(* IEC 61131-3 sources: PLC-IsaVODE/PLC-IsaVODE/samples/plc-programs (part 12) *)

(* ---- 716-TIMER_2.ST ---- *)
FUNCTION UDINT_TO_TIME2:TIME

	VAR_INPUT
		IN :	UDINT;
	END_VAR

	UDINT_TO_TIME2 := DINT_TO_TIME(UDINT_TO_DINT(IN));

END_FUNCTION

FUNCTION_BLOCK T_PLC_MS_block
	VAR_OUTPUT
		T_PLC_MS :	UDINT;
	END_VAR

	VAR_EXTERNAL
		PLC_TICKS_PER_SEC :	INT;
		PLC_SYS_TICK_CNT :	DINT;
	END_VAR

	VAR
		debug :	BOOL;(*Debug-Mode ON / OFF*)
		N :	INT;(*Debug-Faktor*)
		Offset :	UDINT;(*Debug-Offset*)
		temp :	DWORD := DWORD#1;(*Debug-Offset*)
		mode :	BOOL;(*modus*)
		faktor :	UDINT;(*Systemtakt-Faktor*)
		init :	BOOL;
		v_plc_ticks_per_sec :	UDINT;
		base :	UDINT := UDINT#1000;
	END_VAR

	IF init = FALSE THEN
		v_plc_ticks_per_sec := INT_TO_UDINT(PLC_TICKS_PER_SEC);
		IF v_plc_ticks_per_sec = UDINT#1024 THEN
			faktor := UDINT#1;
			mode := FALSE;
		ELSIF v_plc_ticks_per_sec > UDINT#0 THEN
			IF v_plc_ticks_per_sec <= base THEN
				faktor := base / v_plc_ticks_per_sec;
				mode := FALSE;
			ELSE
				faktor := v_plc_ticks_per_sec / base;
				mode := TRUE;
			END_IF;
		ELSE
			faktor := UDINT#1;
		END_IF;
		init := TRUE;
	END_IF;

	IF mode THEN
		T_PLC_MS := DINT_TO_UDINT(PLC_SYS_TICK_CNT) / faktor;
	ELSE
		T_PLC_MS := DINT_TO_UDINT(PLC_SYS_TICK_CNT) * faktor;
	END_IF;

	IF debug THEN
		T_PLC_MS := (DWORD_TO_UDINT(SHL(UDINT_TO_DWORD(T_PLC_MS),N) OR SHL(temp,N)) - UDINT#1) + Offset;
	END_IF;
END_FUNCTION_BLOCK

FUNCTION DAY_OF_WEEK:INT
  VAR_INPUT
    IDATE :	UDINT;
  END_VAR

  DAY_OF_WEEK := UDINT_TO_INT((idate / UDINT#86400 + UDINT#3) MOD UDINT#7) + INT#01;
END_FUNCTION

FUNCTION _BYTE_TO_INT:INT
	VAR_INPUT
		IN :	BYTE;
	END_VAR

	_BYTE_TO_INT := USINT_TO_INT(BYTE_TO_USINT(IN));
END_FUNCTION

FUNCTION LEAP_OF_DATE:BOOL

	VAR_INPUT
		IDATE :	UDINT;
	END_VAR

	LEAP_OF_DATE := SHL(UDINT_TO_DWORD((idate + UDINT#43200) / UDINT#31557600), 30) = DWORD#16#80000000;

END_FUNCTION

FUNCTION DAY_OF_YEAR:INT
	VAR_INPUT
		IDATE :	DATE;
	END_VAR

	DAY_OF_YEAR := UDINT_TO_INT((DATE_TO_UDINT(idate) / UDINT#86400) MOD UDINT#1461);
	IF DAY_OF_YEAR > 729 THEN
		IF DAY_OF_YEAR > 1095 THEN DAY_OF_YEAR := DAY_OF_YEAR - 1095; ELSE DAY_OF_YEAR := DAY_OF_YEAR - 729; END_IF;
	ELSIF DAY_OF_YEAR > 364 THEN
		DAY_OF_YEAR := DAY_OF_YEAR - 364;
	ELSE
		DAY_OF_YEAR := DAY_OF_YEAR + 1;
	END_IF;
END_FUNCTION

FUNCTION DAY_OF_YEAR_UDINT:INT
	VAR_INPUT
		IDATE :	UDINT;
	END_VAR

	DAY_OF_YEAR_UDINT := UDINT_TO_INT((idate / UDINT#86400) MOD UDINT#1461);
	IF DAY_OF_YEAR_UDINT > 729 THEN
		IF DAY_OF_YEAR_UDINT > 1095 THEN DAY_OF_YEAR_UDINT := DAY_OF_YEAR_UDINT - 1095; ELSE DAY_OF_YEAR_UDINT := DAY_OF_YEAR_UDINT - 729; END_IF;
	ELSIF DAY_OF_YEAR_UDINT > 364 THEN
		DAY_OF_YEAR_UDINT := DAY_OF_YEAR_UDINT - 364;
	ELSE
		DAY_OF_YEAR_UDINT := DAY_OF_YEAR_UDINT + 1;
	END_IF;
END_FUNCTION

FUNCTION MONTH_OF_DATE_UDINT:INT

	VAR_INPUT
		IDATE :	UDINT;
	END_VAR

	MONTH_OF_DATE_UDINT := DAY_OF_YEAR_UDINT(idate);
	IF MONTH_OF_DATE_UDINT < 32 THEN
		MONTH_OF_DATE_UDINT := 1;
	ELSIF LEAP_OF_DATE(IDATE) THEN
		MONTH_OF_DATE_UDINT := (MONTH_OF_DATE_UDINT * 53 + 1668) / 1623;
	ELSE
		MONTH_OF_DATE_UDINT := (MONTH_OF_DATE_UDINT * 53 + 1700) / 1620;
	END_IF;

END_FUNCTION

FUNCTION DAY_OF_MONTH:INT
	VAR_INPUT
		IDATE :	UDINT;
	END_VAR

	day_of_month := day_of_year_UDINT(idate);

	IF leap_of_Date(idate) THEN
		CASE day_of_month OF
			32..60	:	day_of_month := day_of_month - 31;
			61..91	:	day_of_month := day_of_month - 60;
			92..121 :	day_of_month := day_of_month - 91;
			122..152:	day_of_month := day_of_month - 121;
			153..182:	day_of_month := day_of_month - 152;
			183..213:	day_of_month := day_of_month - 182;
			214..244:	day_of_month := day_of_month - 213;
			245..274:	day_of_month := day_of_month - 244;
			275..305:	day_of_month := day_of_month - 274;
			306..335:	day_of_month := day_of_month - 305;
			336..366:	day_of_month := day_of_month - 335;
		END_CASE;
	ELSE
		CASE day_of_month OF
			32..59	:	day_of_month := day_of_month - 31;
			60..90	:	day_of_month := day_of_month - 59;
			91..120 :	day_of_month := day_of_month - 90;
			121..151:	day_of_month := day_of_month - 120;
			152..181:	day_of_month := day_of_month - 151;
			182..212:	day_of_month := day_of_month - 181;
			213..243:	day_of_month := day_of_month - 212;
			244..273:	day_of_month := day_of_month - 243;
			274..304:	day_of_month := day_of_month - 273;
			305..334:	day_of_month := day_of_month - 304;
			335..365:	day_of_month := day_of_month - 334;
		END_CASE;
	END_IF;

END_FUNCTION

FUNCTION MONTH_OF_DATE:INT

	VAR_INPUT
		IDATE :	DATE;
	END_VAR

	MONTH_OF_DATE := DAY_OF_YEAR(idate);
	IF MONTH_OF_DATE < 32 THEN
		MONTH_OF_DATE := 1;
	ELSIF LEAP_OF_DATE(DATE_TO_UDINT(IDATE)) THEN
		MONTH_OF_DATE := (MONTH_OF_DATE * 53 + 1668) / 1623;
	ELSE
		MONTH_OF_DATE := (MONTH_OF_DATE * 53 + 1700) / 1620;
	END_IF;

END_FUNCTION

FUNCTION TIME_TO_UDINT2:UDINT
	VAR_INPUT
		X :	TIME;
	END_VAR

	TIME_TO_UDINT2 := DINT_TO_UDINT(TIME_TO_DINT(X));
END_FUNCTION

FUNCTION DT_TO_TOD2:UDINT
	VAR_INPUT
		IN :	UDINT;
	END_VAR

	DT_TO_TOD2 := (IN MOD UDINT#86400) * UDINT#1000;
END_FUNCTION

FUNCTION _DT_TO_DATE_B:UDINT

	VAR_INPUT
		_INN :	UDINT;
	END_VAR

	_DT_TO_DATE_B := (_INN / UDINT#86400) * UDINT#86400;
END_FUNCTION

FUNCTION_BLOCK TIMER_2_Block

	VAR_INPUT
		DT_IN :	UDINT;
		START :	UDINT;
		DURATION :	TIME;
		MODE :	BYTE;
		HOLIDAY :	BOOL;
	END_VAR

	VAR_OUTPUT
		Q :	BOOL;
	END_VAR

	VAR
		last_check :	TIME := T#0s;
		dat :	UDINT;
		daytime :	UDINT;
		activation :	TIME;
		tx :	TIME;
		enabled :	BOOL;
		wday :	INT;
		init :	BOOL;
	END_VAR

	VAR RETAIN
		run_date :	UDINT;
	END_VAR

	VAR
		T_PLC_MS :	T_PLC_MS_Block;
	END_VAR

	T_PLC_MS();
	tx:= UDINT_TO_TIME(T_PLC_MS.T_PLC_MS);

	IF NOT init THEN
		init := TRUE;
		last_check := tx - t#100ms;
	END_IF;

	IF tx - last_check < T#100ms THEN RETURN; END_IF;

	dat := _DT_TO_DATE_B(dt_in);
	daytime := DT_TO_TOD2(dt_in);
	wday := DAY_OF_WEEK(dat);

	CASE _BYTE_TO_INT(mode) OF
	1..7:
		enabled := wday = _BYTE_TO_INT(mode);
	11:
		enabled := TRUE;
	12..16:
		enabled := (dat / UDINT#86400) MOD (BYTE_TO_UDINT(mode) - UDINT#10) = UDINT#0;
	20:
		enabled := wday <= 5;
	21:
		enabled := wday > 5;
	22:
		enabled := wday <= 5 AND NOT holiday;
	23:
		enabled := wday > 5 OR holiday;
	24:
		enabled := holiday;
	25:
		enabled := DAY_OF_MONTH(dat) = 1;
	26:
		enabled := day_of_month(dat + TIME_TO_UDINT2(t#1d)) = 1;
	27:
		enabled := DAY_OF_MONTH(dat) = 31 AND MONTH_OF_DATE_UDINT(dat) = 12;
	28:
		enabled := DAY_OF_YEAR_UDINT(dat) = 1;
	ELSE
		enabled := FALSE;
	END_CASE;

	IF enabled AND NOT Q AND daytime >= start AND run_date <> dat THEN
		Q := TRUE;
		activation := tx;
		run_date := dat;
	ELSIF Q AND tx - activation >= duration THEN
		Q := FALSE;
	END_IF;
	last_check := Tx;

END_FUNCTION_BLOCK

PROGRAM program0
	VAR
		DT_IN :	UDINT;
		START :	UDINT;
		DURATION :	TIME;
		MODE :	BYTE;
		HOLIDAY :	BOOL;
		Q :	BOOL;

		func_block : TIMER_2_Block;
	END_VAR
	func_block.DT_IN := DT_IN;
	func_block.START := START;
	func_block.DURATION := DURATION ;
	func_block.MODE    := MODE    ;
	func_block.HOLIDAY := HOLIDAY;

	func_block();
	Q  := func_block.Q;
END_PROGRAM

CONFIGURATION Config0
	VAR_GLOBAL
		PLC_TICKS_PER_SEC :	INT;
		PLC_SYS_TICK_CNT :	DINT;
	END_VAR
  	RESOURCE Res0 ON PLC
    	TASK task0(INTERVAL := T#20ms,PRIORITY := 0);
    	PROGRAM instance0 WITH task0 : program0;
  	END_RESOURCE
END_CONFIGURATION

(* ---- 717-SEQUENCE_8.ST ---- *)
FUNCTION UDINT_TO_TIME2:TIME

	VAR_INPUT
		IN :	UDINT;
	END_VAR

	UDINT_TO_TIME2 := DINT_TO_TIME(UDINT_TO_DINT(IN));

END_FUNCTION

FUNCTION_BLOCK T_PLC_MS_block
	VAR_OUTPUT
		T_PLC_MS :	UDINT;
	END_VAR

	VAR_EXTERNAL
		PLC_TICKS_PER_SEC :	INT;
		PLC_SYS_TICK_CNT :	DINT;
	END_VAR

	VAR
		debug :	BOOL;
		N :	INT;
		Offset :	UDINT;
		temp :	DWORD := DWORD#1;
		mode :	BOOL;
		faktor :	UDINT;
		init :	BOOL;
		v_plc_ticks_per_sec :	UDINT;
		base :	UDINT := UDINT#1000;
	END_VAR

	IF init = FALSE THEN
		v_plc_ticks_per_sec := INT_TO_UDINT(PLC_TICKS_PER_SEC);
		IF v_plc_ticks_per_sec = UDINT#1024 THEN
			faktor := UDINT#1;
			mode := FALSE;
		ELSIF v_plc_ticks_per_sec > UDINT#0 THEN
			IF v_plc_ticks_per_sec <= base THEN
				faktor := base / v_plc_ticks_per_sec;
				mode := FALSE;
			ELSE
				faktor := v_plc_ticks_per_sec / base;
				mode := TRUE;
			END_IF;
		ELSE
			faktor := UDINT#1;
		END_IF;
		init := TRUE;
	END_IF;

	IF mode THEN
		T_PLC_MS := DINT_TO_UDINT(PLC_SYS_TICK_CNT) / faktor;
	ELSE
		T_PLC_MS := DINT_TO_UDINT(PLC_SYS_TICK_CNT) * faktor;
	END_IF;

	IF debug THEN
		T_PLC_MS := (DWORD_TO_UDINT(SHL(UDINT_TO_DWORD(T_PLC_MS),N) OR SHL(temp,N)) - UDINT#1) + Offset;
	END_IF;

END_FUNCTION_BLOCK

FUNCTION_BLOCK SEQUENCE_8_Block

	VAR_INPUT
		IN0 :	BOOL := TRUE;
		IN1 :	BOOL := TRUE;
		IN2 :	BOOL := TRUE;
		IN3 :	BOOL := TRUE;
		IN4 :	BOOL := TRUE;
		IN5 :	BOOL := TRUE;
		IN6 :	BOOL := TRUE;
		IN7 :	BOOL := TRUE;
		START :	BOOL;
		RST :	BOOL;
		WAIT0 :	TIME;
		DELAY0 :	TIME;
		WAIT1 :	TIME;
		DELAY1 :	TIME;
		WAIT2 :	TIME;
		DELAY2 :	TIME;
		WAIT3 :	TIME;
		DELAY3 :	TIME;
		WAIT4 :	TIME;
		DELAY4 :	TIME;
		WAIT5 :	TIME;
		DELAY5 :	TIME;
		WAIT6 :	TIME;
		DELAY6 :	TIME;
		WAIT7 :	TIME;
		DELAY7 :	TIME;
		STOP_ON_ERROR :	BOOL;
	END_VAR

	VAR_OUTPUT
		Q0 :	BOOL;
		Q1 :	BOOL;
		Q2 :	BOOL;
		Q3 :	BOOL;
		Q4 :	BOOL;
		Q5 :	BOOL;
		Q6 :	BOOL;
		Q7 :	BOOL;
		QX :	BOOL;
		RUN :	BOOL;
		_STEP :	INT := -1;
		STATUS :	BYTE;
	END_VAR

	VAR
		last :	TIME;
		edge :	BOOL;
		tx :	TIME;
		init :	BOOL;
		T_PLC_MS :	T_PLC_MS_Block;
	END_VAR

	T_PLC_MS();
	tx:= UDINT_TO_TIME(T_PLC_MS.T_PLC_MS);

	IF NOT init THEN
		last := tx;
		init := TRUE;
		status := BYTE#110;
	END_IF;

	IF rst THEN
		_step := -1;
		Q0 := FALSE;
		Q1 := FALSE;
		Q2 := FALSE;
		Q3 := FALSE;
		Q4 := FALSE;
		Q5 := FALSE;
		Q6 := FALSE;
		Q7 := FALSE;
		status := BYTE#110;
		run := FALSE;

	ELSIF start AND NOT edge THEN
		_step := 0;
		last := tx;
		status := BYTE#111;
		Q0 := FALSE;
		Q1 := FALSE;
		Q2 := FALSE;
		Q3 := FALSE;
		Q4 := FALSE;
		Q5 := FALSE;
		Q6 := FALSE;
		Q7 := FALSE;
		run := TRUE;
	END_IF;
	edge := start;

	IF status > BYTE#0 AND status < BYTE#100 AND stop_on_error THEN RETURN; END_IF;

	IF run AND _step = 0 THEN
		IF NOT q0 AND in0 AND tx - last <= wait0 THEN
			Q0 := TRUE;
			last := tx;
		ELSIF NOT q0 AND tx - last > wait0 THEN
			status := BYTE#1;
			run := FALSE;
		ELSIF q0 AND tx - last >= delay0 THEN
			_step := 1;
			last := tx;
		END_IF;
	END_IF;
	IF run AND _step = 1 THEN
		IF NOT q1 AND in1 AND tx - last <= wait1 THEN
			Q0 := FALSE;
			Q1 := TRUE;
			last := tx;
		ELSIF NOT q1 AND Tx - last > wait1 THEN
			status := BYTE#2;
			q0 := FALSE;
			run := FALSE;
		ELSIF q1 AND tx - last >= delay1 THEN
			_step := 2;
			last := tx;
		END_IF;
	END_IF;
	IF run AND _step = 2 THEN
		IF NOT q2 AND in2 AND tx - last <= wait2 THEN
			Q1 := FALSE;
			Q2 := TRUE;
			last := tx;
		ELSIF NOT q2 AND Tx - last > wait2 THEN
			status := BYTE#3;
			q1 := FALSE;
			run := FALSE;
		ELSIF q2 AND tx - last >= delay2 THEN
			_step := 3;
			last := tx;
		END_IF;
	END_IF;
	IF run AND _step = 3 THEN
		IF NOT q3 AND in3 AND tx - last <= wait3 THEN
			Q2 := FALSE;
			Q3 := TRUE;
			last := tx;
		ELSIF NOT q3 AND Tx - last > wait3 THEN
			status := BYTE#4;
			q2 := FALSE;
			run := FALSE;
		ELSIF q3 AND tx - last >= delay3 THEN
			_step := 4;
			last := tx;
		END_IF;
	END_IF;
	IF run AND _step = 4 THEN
		IF NOT q4 AND in4 AND tx - last <= wait4 THEN
			Q3 := FALSE;
			Q4 := TRUE;
			last := tx;
		ELSIF NOT q4 AND Tx - last > wait4 THEN
			status := BYTE#5;
			q3 := FALSE;
			run := FALSE;
		ELSIF q4 AND tx - last >= delay4 THEN
			_step := 5;
			last := tx;
		END_IF;
	END_IF;
	IF run AND _step = 5 THEN
		IF NOT q5 AND in5 AND tx - last <= wait5 THEN
			Q4 := FALSE;
			Q5 := TRUE;
			last := tx;
		ELSIF NOT q5 AND Tx - last > wait5 THEN
			status := BYTE#6;
			q4 := FALSE;
			run := FALSE;
		ELSIF q5 AND tx - last >= delay5 THEN
			_step := 6;
			last := tx;
		END_IF;
	END_IF;
	IF run AND _step = 6 THEN
		IF NOT q6 AND in6 AND tx - last <= wait6 THEN
			Q5 := FALSE;
			Q6 := TRUE;
			last := tx;
		ELSIF NOT q6 AND Tx - last > wait6 THEN
			status := BYTE#7;
			q5 := FALSE;
			run := FALSE;
		ELSIF q6 AND tx - last >= delay6 THEN
			_step := 7;
			last := tx;
		END_IF;
	END_IF;
	IF run AND _step = 7 THEN
		IF NOT q7 AND in7 AND tx - last <= wait7 THEN
			Q6 := FALSE;
			Q7 := TRUE;
			last := tx;
		ELSIF NOT q7 AND Tx - last > wait7 THEN
			status := BYTE#8;
			q6 := FALSE;
			run := FALSE;
		ELSIF q7 AND tx - last >= delay7 THEN
			_step := -1;
			Q7 := FALSE;
			Run := FALSE;
			status := BYTE#110;
		END_IF;
	END_IF;
	QX := q0 OR q1 OR q2 OR q3 OR q4 OR q5 OR q6 OR q7;

END_FUNCTION_BLOCK

PROGRAM program0

	VAR
		IN0 :	BOOL := TRUE;
		IN1 :	BOOL := TRUE;
		IN2 :	BOOL := TRUE;
		IN3 :	BOOL := TRUE;
		IN4 :	BOOL := TRUE;
		IN5 :	BOOL := TRUE;
		IN6 :	BOOL := TRUE;
		IN7 :	BOOL := TRUE;
		START :	BOOL;
		RST :	BOOL;
		WAIT0 :	TIME;
		DELAY0 :	TIME;
		WAIT1 :	TIME;
		DELAY1 :	TIME;
		WAIT2 :	TIME;
		DELAY2 :	TIME;
		WAIT3 :	TIME;
		DELAY3 :	TIME;
		WAIT4 :	TIME;
		DELAY4 :	TIME;
		WAIT5 :	TIME;
		DELAY5 :	TIME;
		WAIT6 :	TIME;
		DELAY6 :	TIME;
		WAIT7 :	TIME;
		DELAY7 :	TIME;
		STOP_ON_ERROR :	BOOL;
		Q0 :	BOOL;
		Q1 :	BOOL;
		Q2 :	BOOL;
		Q3 :	BOOL;
		Q4 :	BOOL;
		Q5 :	BOOL;
		Q6 :	BOOL;
		Q7 :	BOOL;
		QX :	BOOL;
		RUN :	BOOL;
		_STEP :	INT := -1;
		STATUS :	BYTE;
		func_block : SEQUENCE_8_Block;
  	END_VAR
	func_block.IN0  :=IN0;
	func_block.IN1  :=IN1;
	func_block.IN2  :=IN2;
	func_block.IN3  :=IN3;
	func_block.IN4  :=IN4;
	func_block.IN5  :=IN5;
	func_block.IN6  :=IN6;
	func_block.IN7  :=IN7;
	func_block.START  :=START;
	func_block.RST  :=RST;
	func_block.WAIT0  :=WAIT0;
	func_block.DELAY0  :=DELAY0;
	func_block.WAIT1:=WAIT1;
	func_block.DELAY1:=DELAY1;
	func_block.WAIT2  :=WAIT2;
	func_block.DELAY2  :=DELAY2;
	func_block.WAIT3  :=WAIT3;
	func_block.DELAY3  :=DELAY3;
	func_block.DELAY1:=DELAY1;
	func_block.WAIT2  :=WAIT2;
	func_block.DELAY2  :=DELAY2;
	func_block.WAIT3  :=WAIT3;
	func_block.DELAY3  :=DELAY3;
	func_block.WAIT4:=WAIT4;
	func_block.DELAY4  :=DELAY4;
	func_block.WAIT5  :=WAIT5;
	func_block.DELAY5  :=DELAY5;
	func_block.WAIT6  :=WAIT6;
	func_block.DELAY6  :=DELAY6;
	func_block.WAIT7  :=WAIT7;
	func_block.DELAY7  :=DELAY7;
	func_block.STOP_ON_ERROR  :=STOP_ON_ERROR;
	func_block();
	Q0 := func_block.Q0;
	Q1 := func_block.Q1;
	Q2 := func_block.Q2;
	Q3 := func_block.Q3;
	Q4 := func_block.Q4;
	Q5 := func_block.Q5;
	Q6 := func_block.Q6;
	Q7 := func_block.Q7;
	QX := func_block.QX;
	RUN := func_block.RUN;
	_STEP := func_block._STEP;
	STATUS := func_block.STATUS;

END_PROGRAM

CONFIGURATION Config0

	VAR_GLOBAL
		PLC_TICKS_PER_SEC :	INT;
		PLC_SYS_TICK_CNT :	DINT;
	END_VAR

	RESOURCE Res0 ON PLC
		TASK task0(INTERVAL := T#20ms,PRIORITY := 0);
		PROGRAM instance0 WITH task0 : program0;
	END_RESOURCE

END_CONFIGURATION

(* ---- 718-BLIND_INPUT.ST ---- *)
FUNCTION UDINT_TO_TIME2:TIME

	VAR_INPUT
		IN :	UDINT;
	END_VAR

	UDINT_TO_TIME2 := DINT_TO_TIME(UDINT_TO_DINT(IN));

END_FUNCTION

FUNCTION_BLOCK T_PLC_MS_block
	VAR_OUTPUT
		T_PLC_MS :	UDINT;
	END_VAR

	VAR_EXTERNAL
		PLC_TICKS_PER_SEC :	INT;
		PLC_SYS_TICK_CNT :	DINT;
	END_VAR

	VAR
		debug :	BOOL;(*Debug-Mode ON / OFF*)
		N :	INT;(*Debug-Faktor*)
		Offset :	UDINT;(*Debug-Offset*)
		temp :	DWORD := DWORD#1;(*Debug-Offset*)
		mode :	BOOL;(*modus*)
		faktor :	UDINT;(*Systemtakt-Faktor*)
		init :	BOOL;
		v_plc_ticks_per_sec :	UDINT;
		base :	UDINT := UDINT#1000;
	END_VAR

	IF init = FALSE THEN
		v_plc_ticks_per_sec := INT_TO_UDINT(PLC_TICKS_PER_SEC);
		IF v_plc_ticks_per_sec = UDINT#1024 THEN
			faktor := UDINT#1;
			mode := FALSE;
		ELSIF v_plc_ticks_per_sec > UDINT#0 THEN
			IF v_plc_ticks_per_sec <= base THEN
				faktor := base / v_plc_ticks_per_sec;
				mode := FALSE;
			ELSE
				faktor := v_plc_ticks_per_sec / base;
				mode := TRUE;
			END_IF;
		ELSE
			faktor := UDINT#1;
		END_IF;
		init := TRUE;
	END_IF;

	IF mode THEN
		T_PLC_MS := DINT_TO_UDINT(PLC_SYS_TICK_CNT) / faktor;
	ELSE
		T_PLC_MS := DINT_TO_UDINT(PLC_SYS_TICK_CNT) * faktor;
	END_IF;

	IF debug THEN
		T_PLC_MS := (DWORD_TO_UDINT(SHL(UDINT_TO_DWORD(T_PLC_MS),N) OR SHL(temp,N)) - UDINT#1) + Offset;
	END_IF;

END_FUNCTION_BLOCK

FUNCTION_BLOCK CLICK_MODE_Block

	VAR_INPUT
		IN :	BOOL;
		T_LONG :	TIME := T#500ms;
	END_VAR

	VAR_OUTPUT
		SINGLE_ :	BOOL;
		DOUBLE :	BOOL;
		LONG :	BOOL;
		TP_LONG :	BOOL;
	END_VAR

	VAR
		Timer :	TP;
		cnt :	INT;
		last :	BOOL;
	END_VAR

	timer(in := IN, PT := T_LONG);
	single := FALSE;
	double := FALSE;

	IF timer.Q THEN
		IF NOT in AND last THEN	cnt := cnt + 1; END_IF;
	ELSE
		CASE cnt OF
			1 : single := TRUE;
			2 : double := TRUE;
		END_CASE;
		cnt := 0;
	END_IF;
	last := in;
	TP_LONG := NOT timer.Q AND (NOT LONG) AND IN;
	LONG := NOT timer.Q AND in;

END_FUNCTION_BLOCK

FUNCTION _BYTE_TO_INT:INT
	VAR_INPUT
		IN :	BYTE;
	END_VAR

	_BYTE_TO_INT := USINT_TO_INT(BYTE_TO_USINT(IN));
END_FUNCTION

FUNCTION_BLOCK BLIND_INPUT_Block

	VAR_INPUT
		POS :	BYTE;
		ANG :	BYTE;
		S1 :	BOOL;
		S2 :	BOOL;
		IN :	BOOL;
		PI :	BYTE;
		AI :	BYTE;
		SINGLE_SWITCH :	BOOL;
		CLICK_EN :	BOOL := TRUE;
		CLICK_TIME :	TIME := T#500ms;
		MAX_RUNTIME :	TIME := T#60s;
		MANUAL_TIMEOUT :	TIME := T#1h;
		DEBOUNCE_TIME :	TIME := T#20ms;
		DBL_CLK1 :	BOOL := FALSE;
		DBL_POS1 :	BYTE;
		DBL_ANG1 :	BYTE;
		DBL_CLK2 :	BOOL := FALSE;
		DBL_POS2 :	BYTE := BYTE#255;
		DBL_ANG2 :	BYTE := BYTE#255;
		D1_TOGGLE :	BOOL := TRUE;
		D2_TOGGLE :	BOOL := TRUE;
		MASTER_MODE :	BOOL;
	END_VAR

	VAR_OUTPUT
		QU :	BOOL := TRUE;
		QD :	BOOL := TRUE;
		STATUS :	BYTE;
		PO :	BYTE := BYTE#255;
		AO :	BYTE := BYTE#255;
		D1 :	BOOL;
		D2 :	BOOL;
	END_VAR

	VAR
		s1e :	TOF;
		s2e :	TOF;
		s1d :	CLICK_MODE_Block;
		s2d :	CLICK_MODE_Block;
		dir :	BOOL;
		tx :	TIME;
		last :	TIME;
		T_PLC_MS :	T_PLC_MS_Block;
	END_VAR

	T_PLC_MS();
	tx:= UDINT_TO_TIME(T_PLC_MS.T_PLC_MS);

	s1e(in := S1, pt := DEBOUNCE_TIME);
	s2e(in := S2, pt := DEBOUNCE_TIME);
	s1d(in := (s1e.Q AND NOT SINGLE_SWITCH) OR (s1e.Q AND SINGLE_SWITCH AND dir), t_long := CLICK_TIME);
	s2d(in := (s2e.Q AND NOT SINGLE_SWITCH) OR (s1e.Q AND SINGLE_SWITCH AND NOT dir), t_long := CLICK_TIME);

	IF NOT d1_toggle THEN d1 := FALSE; END_IF;
	IF NOT d2_toggle THEN d2 := FALSE; END_IF;

	IF (s1d.LONG AND s2d.LONG) OR (status = BYTE#139) THEN
	status := BYTE#139;
	IF NOT (s1d.LONG OR s2d.LONG)  THEN status := BYTE#130; END_IF;
	ELSIF s1d.tp_LONG THEN
		status := BYTE#132;
	ELSIF s2d.tp_LONG THEN
		status := BYTE#133;
	ELSIF  s1d.SINGLE_ THEN
		IF click_en THEN
			IF QU XOR QD THEN
				status := BYTE#131;
			ELSE
				status := BYTE#134;
				last := tx;
				dir := NOT dir;
			END_IF;
		END_IF;
	ELSIF  s2d.SINGLE_ THEN
		IF click_en THEN
			IF QU XOR QD THEN
				status := BYTE#131;
			ELSE
				status := BYTE#135;
				last := tx;
				dir := NOT dir;
			END_IF;
		END_IF;
	ELSIF in THEN
		status := BYTE#136;
		last := tx;
	ELSIF s1d.DOUBLE THEN
		IF dbl_clk1 THEN
			status := BYTE#137;
			last := tx;
		ELSE
			D1 := NOT D1;
		END_IF;
	ELSIF s2d.DOUBLE THEN
		IF dbl_clk2 THEN
			status := BYTE#138;
			last := tx;
		ELSE
			IF single_switch THEN D1 := NOT D1; ELSE D2 := NOT D2; END_IF;
		END_IF;
	END_IF;

	CASE _BYTE_TO_INT(status) OF
		0:
				status := BYTE#130;

		130:
				IF NOT master_mode THEN
					PO := POS;
					AO := ANG;
				END_IF;
				QU := TRUE;
				QD := TRUE;

		131:
				QU := FALSE;
				QD := FALSE;
				PO := POS;
				AO := ANG;
				IF tx - last >= manual_timeout THEN
					status := BYTE#130;
				END_IF;

		132:
				QU := TRUE;
				QD := FALSE;
				PO := POS; AO := ANG;
				last := tx;
				IF NOT s1d.LONG THEN status := BYTE#131; dir := NOT dir; END_IF;

		133:
				QU := FALSE;
				QD := TRUE;
				PO := POS; AO := ANG;
				last := tx;
				IF NOT s2d.LONG THEN	status := BYTE#131; dir := NOT dir; END_IF;

		134:
				QU := TRUE;
				QD := FALSE;
				PO := POS; AO := ANG;
				IF tx - last >= max_runtime THEN status := BYTE#131; END_IF;

		135:
				QU := FALSE;
				QD := TRUE;
				PO := POS; AO := ANG;
				IF tx - last >= max_runtime THEN status := BYTE#131;	END_IF;

		136:
				QU := TRUE;
				QD := TRUE;
				PO := PI; AO := AI;
				IF tx-last >= max_runtime THEN status := BYTE#130; END_IF;

		137:
				QU := TRUE;
				QD := TRUE;
				PO := DBL_POS1;
				AO := DBL_ANG1;
				IF tx - last >= max_runtime THEN status := BYTE#131; END_IF;

		138:
				QU := TRUE;
				QD := TRUE;
				PO := DBL_POS2;
				AO := DBL_ANG2;
				IF tx - last >= max_runtime THEN status := BYTE#131; END_IF;

		139:
				QU := FALSE;
				QD := FALSE;
				PO := POS;
				AO := ANG;

	END_CASE;

END_FUNCTION_BLOCK

PROGRAM program0
	VAR
		POS :	BYTE;
		ANG :	BYTE;
		S1 :	BOOL;
		S2 :	BOOL;
		IN :	BOOL;
		PI :	BYTE;
		AI :	BYTE;
		SINGLE_SWITCH :	BOOL;
		CLICK_EN :	BOOL := TRUE;
		CLICK_TIME :	TIME := T#500ms;
		MAX_RUNTIME :	TIME := T#60s;
		MANUAL_TIMEOUT :	TIME := T#1h;
		DEBOUNCE_TIME :	TIME := T#20ms;
		DBL_CLK1 :	BOOL := FALSE;
		DBL_POS1 :	BYTE;
		DBL_ANG1 :	BYTE;
		DBL_CLK2 :	BOOL := FALSE;
		DBL_POS2 :	BYTE := BYTE#255;
		DBL_ANG2 :	BYTE := BYTE#255;
		D1_TOGGLE :	BOOL := TRUE;
		D2_TOGGLE :	BOOL := TRUE;
		MASTER_MODE :	BOOL;
		QU :	BOOL := TRUE;
		QD :	BOOL := TRUE;
		STATUS :	BYTE;
		PO :	BYTE := BYTE#255;
		AO :	BYTE := BYTE#255;
		D1 :	BOOL;
		D2 :	BOOL;
		func_block : BLIND_INPUT_Block;
	END_VAR
	func_block.POS := POS;
	func_block.ANG := ANG;
	func_block.S1 := S1 ;
	func_block.S2 := S2;
	func_block.IN := IN;
	func_block.PI := PI;
	func_block.AI := AI;
	func_block.SINGLE_SWITCH := SINGLE_SWITCH;
	func_block.CLICK_EN := CLICK_EN ;
	func_block.CLICK_TIME := CLICK_TIME;
	func_block.MAX_RUNTIME := MAX_RUNTIME;
	func_block.MANUAL_TIMEOUT := MANUAL_TIMEOUT;
	func_block.DEBOUNCE_TIME := DEBOUNCE_TIME;
	func_block.DBL_CLK1 := DBL_CLK1;
	func_block.DBL_POS1 := DBL_POS1 ;
	func_block.DBL_ANG1 := DBL_ANG1;
	func_block.DBL_CLK2 := DBL_CLK2;
	func_block.DBL_POS2 := DBL_POS2;
	func_block.DBL_ANG2 := DBL_ANG2;
	func_block.D1_TOGGLE := D1_TOGGLE ;
	func_block.D2_TOGGLE := D2_TOGGLE;
	func_block.MASTER_MODE := MASTER_MODE;
	func_block();
	QU  := func_block.QU;
	QD  := func_block.QD;
	STATUS  := func_block.STATUS;
	PO  := func_block.PO;
	AO  := func_block.AO;
	D1  := func_block.D1;
	D2  := func_block.D2;
END_PROGRAM

CONFIGURATION Config0
	VAR_GLOBAL
		PLC_TICKS_PER_SEC :	INT;
		PLC_SYS_TICK_CNT :	DINT;
	END_VAR
  	RESOURCE Res0 ON PLC
    	TASK task0(INTERVAL := T#20ms,PRIORITY := 0);
    	PROGRAM instance0 WITH task0 : program0;
  	END_RESOURCE
END_CONFIGURATION

(* ---- 719-TN_INPUT_MENU_POPUP.ST ---- *)
FUNCTION_BLOCK TN_INPUT_MENU_POPUP

  VAR
    FB_TN_SC_AREA_SAVE :	TN_SC_AREA_SAVE;
    FB_TN_SC_AREA_RESTORE :	TN_SC_AREA_RESTORE;
    FB_TN_SC_LINE :	TN_SC_LINE;
    FB_TN_SC_ADD_SHADOW :	TN_SC_ADD_SHADOW;
    FB_TN_SC_BOX :	TN_SC_BOX;
    FB_TN_SC_WRITE_C :	TN_SC_WRITE_C;
    ELEMENT_COUNT :	ELEMENT_COUNT;
    ELEMENT_GET :	ELEMENT_GET;
  END_VAR

  VAR
    in_ROW :	INT;
    in_ROWS :	INT;
    in_COL :	INT;
    in_COLS :	INT;
    in_index :	INT;
    in_Count :	INT;
    in_Scroll_Offset :	INT;
    by_ATTR :	BYTE;
  END_VAR

  VAR_IN_OUT
    Xus_TN_MENU_POPUP :	us_TN_MENU_POPUP;
    Xus_TN_SCREEN :	us_TN_SCREEN;
  END_VAR

  IF (Xus_TN_MENU_POPUP.bo_Activ = FALSE) AND (Xus_TN_MENU_POPUP.bo_Create = TRUE) THEN
    Xus_TN_MENU_POPUP.bo_Activ         := TRUE;
    Xus_TN_MENU_POPUP.bo_Create        := FALSE;
    Xus_TN_MENU_POPUP.bo_Destroy       := FALSE;
    Xus_TN_MENU_POPUP.bo_Update        := TRUE;

    ELEMENT_COUNT(ELEMENT:=Xus_TN_MENU_POPUP.st_Menu_Text,SEP:=BYTE#35);
    Xus_TN_MENU_POPUP.st_Menu_Text:=ELEMENT_COUNT.ELEMENT;
    Xus_TN_MENU_POPUP.in_Menu_E_Count:=ELEMENT_COUNT.ELEMENT_COUNT;

    Xus_TN_MENU_POPUP.in_Rows := Xus_TN_MENU_POPUP.in_Menu_E_Count;

    Xus_TN_MENU_POPUP.in_Cols := INT#00;

    FOR in_Count := INT#01 TO Xus_TN_MENU_POPUP.in_Rows DO;

      ELEMENT_GET(ELEMENT:=Xus_TN_MENU_POPUP.st_Menu_Text,SEP:=BYTE#35,POS:=in_Count-1);
      Xus_TN_MENU_POPUP.st_Menu_Text:=ELEMENT_GET.ELEMENT;
      Xus_TN_MENU_POPUP.in_Cols:=MAX_INT(LEN(ELEMENT_GET.ELEMENT_GET),Xus_TN_MENU_POPUP.in_Cols);

    END_FOR;

    IF (Xus_TN_MENU_POPUP.in_X + Xus_TN_MENU_POPUP.in_Cols) > INT#75 THEN
      Xus_TN_MENU_POPUP.in_X := INT#79 - Xus_TN_MENU_POPUP.in_Cols - INT#04;
    END_IF;

    IF (Xus_TN_MENU_POPUP.in_Y + Xus_TN_MENU_POPUP.in_ROWS) > INT#21 THEN
      Xus_TN_MENU_POPUP.in_Y := INT#23 - Xus_TN_MENU_POPUP.in_ROWS - INT#2;
    END_IF;

    Xus_TN_SCREEN.bo_Modal_Dialog := TRUE;

    FB_TN_SC_AREA_SAVE.Iin_X1        := Xus_TN_MENU_POPUP.in_X;
    FB_TN_SC_AREA_SAVE.Iin_Y1        := Xus_TN_MENU_POPUP.in_Y;
    FB_TN_SC_AREA_SAVE.Iin_X2        := Xus_TN_MENU_POPUP.in_X + Xus_TN_MENU_POPUP.in_Cols + INT#04;
    FB_TN_SC_AREA_SAVE.Iin_Y2        := Xus_TN_MENU_POPUP.in_Y + Xus_TN_MENU_POPUP.in_Rows + INT#02;
    FB_TN_SC_AREA_SAVE.Xus_TN_SCREEN := Xus_TN_SCREEN;
    FB_TN_SC_AREA_SAVE();
    Xus_TN_SCREEN := FB_TN_SC_AREA_SAVE.Xus_TN_SCREEN;

    FB_TN_SC_BOX.Iin_X1        := Xus_TN_MENU_POPUP.in_X;
    FB_TN_SC_BOX.Iin_Y1        := Xus_TN_MENU_POPUP.in_Y;
    FB_TN_SC_BOX.Iin_X2        := Xus_TN_MENU_POPUP.in_X + Xus_TN_MENU_POPUP.in_Cols + INT#03;
    FB_TN_SC_BOX.Iin_Y2        := Xus_TN_MENU_POPUP.in_Y + Xus_TN_MENU_POPUP.in_Rows + INT#01;
    FB_TN_SC_BOX.Iby_FILL      := BYTE#32;
    FB_TN_SC_BOX.Iin_BORDER    := INT#01;
    FB_TN_SC_BOX.Iby_ATTR      := Xus_TN_MENU_POPUP.by_Attr_oF;
    FB_TN_SC_BOX.Xus_TN_SCREEN := Xus_TN_SCREEN;
    FB_TN_SC_BOX();
    Xus_TN_SCREEN := FB_TN_SC_BOX.Xus_TN_SCREEN;

    FB_TN_SC_ADD_SHADOW.Iin_X1        := Xus_TN_MENU_POPUP.in_X + INT#1;
    FB_TN_SC_ADD_SHADOW.Iin_Y1        := Xus_TN_MENU_POPUP.in_Y + INT#1;
    FB_TN_SC_ADD_SHADOW.Iin_X2        := Xus_TN_MENU_POPUP.in_X + Xus_TN_MENU_POPUP.in_Cols + INT#04;
    FB_TN_SC_ADD_SHADOW.Iin_Y2        := Xus_TN_MENU_POPUP.in_Y + Xus_TN_MENU_POPUP.in_Rows + INT#02;
    FB_TN_SC_ADD_SHADOW.Iin_OPTION    := INT#00;
    FB_TN_SC_ADD_SHADOW.Xus_TN_SCREEN := Xus_TN_SCREEN;
    FB_TN_SC_ADD_SHADOW();
    Xus_TN_SCREEN := FB_TN_SC_ADD_SHADOW.Xus_TN_SCREEN;

    in_COL  := Xus_TN_MENU_POPUP.in_X;
    in_ROW  := Xus_TN_MENU_POPUP.in_Y;
    in_ROWS := Xus_TN_MENU_POPUP.in_Rows;
    in_COLS := Xus_TN_MENU_POPUP.in_Cols;

    in_COLS := in_COLS + INT#02;

    FOR in_Count := INT#01 TO Xus_TN_MENU_POPUP.in_Menu_E_Count DO;
      in_ROW := in_ROW + INT#01;

      ELEMENT_GET(ELEMENT:=Xus_TN_MENU_POPUP.st_Menu_Text,SEP:=BYTE#35,POS:=in_Count-1);
    Xus_TN_MENU_POPUP.st_Menu_Text:=ELEMENT_GET.ELEMENT;

      IF EQ_STRING(ELEMENT_GET.ELEMENT_GET,'-') THEN

        FB_TN_SC_LINE.Iin_Y1			:= in_ROW;
        FB_TN_SC_LINE.Iin_X1			:= in_COL;
        FB_TN_SC_LINE.Iin_Y2			:= in_ROW;
        FB_TN_SC_LINE.Iin_X2			:= in_COL + in_COLS + INT#01;
        FB_TN_SC_LINE.Iby_ATTR		:= Xus_TN_MENU_POPUP.by_Attr_oF;
        FB_TN_SC_LINE.Iby_BORDER		:= BYTE#01;
        FB_TN_SC_LINE.Xus_TN_SCREEN	:= Xus_TN_SCREEN;
        FB_TN_SC_LINE();
        Xus_TN_SCREEN := FB_TN_SC_LINE.Xus_TN_SCREEN;

      END_IF;
    END_FOR;
  END_IF;

  IF (Xus_TN_MENU_POPUP.bo_Activ = TRUE) THEN

    CASE _BYTE_TO_INT(Xus_TN_MENU_POPUP.by_Input_Exten_Code) OF

    65:
      in_Scroll_Offset := INT#-1;
      Xus_TN_MENU_POPUP.bo_Update := TRUE;

    66:
      in_Scroll_Offset := INT#1;
      Xus_TN_MENU_POPUP.bo_Update := TRUE;

    13:
      Xus_TN_MENU_POPUP.bo_Destroy := TRUE;

    27:
      Xus_TN_MENU_POPUP.bo_Destroy := TRUE;
      Xus_TN_MENU_POPUP.in_Cur_Item := INT#00;

    67..68:
      Xus_TN_MENU_POPUP.bo_Destroy := TRUE;
      Xus_TN_MENU_POPUP.in_Cur_Item := INT#00;

    END_CASE;

  END_IF;

  IF (Xus_TN_MENU_POPUP.bo_Activ = TRUE) AND (Xus_TN_MENU_POPUP.bo_Update = TRUE) THEN

    Xus_TN_MENU_POPUP.bo_Update := FALSE;

    in_index := Xus_TN_MENU_POPUP.in_Cur_Item;

    IF (in_index < INT#01) OR (in_index > Xus_TN_MENU_POPUP.in_Menu_E_Count) THEN
      in_Scroll_Offset := INT#01;
      in_index := Xus_TN_MENU_POPUP.in_Menu_E_Count;
    END_IF;

    ELEMENT_GET(ELEMENT:=Xus_TN_MENU_POPUP.st_Menu_Text,SEP:=BYTE#35,POS:=in_index-1);
    Xus_TN_MENU_POPUP.st_Menu_Text:=ELEMENT_GET.ELEMENT;

    IF EQ_STRING(ELEMENT_GET.ELEMENT_GET,'-') THEN
      in_Scroll_Offset := INT#01;
    END_IF;

    IF in_Scroll_Offset <> INT#00 THEN

      FOR in_Count := INT#01 TO Xus_TN_MENU_POPUP.in_Menu_E_Count DO;

        in_index:=INC2(in_index,in_Scroll_Offset,1,Xus_TN_MENU_POPUP.in_Menu_E_Count);

        ELEMENT_GET(ELEMENT:=Xus_TN_MENU_POPUP.st_Menu_Text,SEP:=BYTE#35,POS:=in_index-1);
        Xus_TN_MENU_POPUP.st_Menu_Text:=ELEMENT_GET.ELEMENT;

        IF NE_STRING(ELEMENT_GET.ELEMENT_GET,'-') THEN
          EXIT;
        END_IF;

      END_FOR;
    END_IF;

    Xus_TN_MENU_POPUP.in_Cur_Item := in_index;
    in_Scroll_Offset := INT#00;

    in_COL  := Xus_TN_MENU_POPUP.in_X;
    in_ROW  := Xus_TN_MENU_POPUP.in_Y;
    in_ROWS := Xus_TN_MENU_POPUP.in_Rows;
    in_COLS := Xus_TN_MENU_POPUP.in_Cols;

    in_COLS := in_COLS + INT#02;

    FOR in_Count := INT#01 TO Xus_TN_MENU_POPUP.in_Menu_E_Count DO;

      in_ROW := in_ROW + INT#01;

      IF in_Count = Xus_TN_MENU_POPUP.in_Cur_Item THEN
        by_ATTR := Xus_TN_MENU_POPUP.by_Attr_mF;
      ELSE
        by_ATTR := Xus_TN_MENU_POPUP.by_Attr_oF;
      END_IF;

      ELEMENT_GET(ELEMENT:=Xus_TN_MENU_POPUP.st_Menu_Text,SEP:=BYTE#35,POS:=in_Count-1);
      Xus_TN_MENU_POPUP.st_Menu_Text:=ELEMENT_GET.ELEMENT;

      IF NE_STRING(ELEMENT_GET.ELEMENT_GET,'-') THEN

        FB_TN_SC_WRITE_C.Iin_Y         := in_ROW;
        FB_TN_SC_WRITE_C.Iin_X         := in_COL + INT#01;
        FB_TN_SC_WRITE_C.Iby_ATTR      := by_ATTR;
        FB_TN_SC_WRITE_C.Iin_LENGTH    := in_COLS;
        FB_TN_SC_WRITE_C.Iin_OPTION    := INT#02;
        FB_TN_SC_WRITE_C.Ist_STRING    := ELEMENT_GET.ELEMENT_GET;
        FB_TN_SC_WRITE_C.Xus_TN_SCREEN := Xus_TN_SCREEN;
        FB_TN_SC_WRITE_C();
        Xus_TN_SCREEN := FB_TN_SC_WRITE_C.Xus_TN_SCREEN;

      END_IF;
    END_FOR;
  END_IF;

  IF (Xus_TN_MENU_POPUP.bo_Activ = TRUE) AND (Xus_TN_MENU_POPUP.bo_Destroy = TRUE) THEN

    Xus_TN_MENU_POPUP.bo_Destroy := FALSE;
    Xus_TN_MENU_POPUP.bo_Activ   := FALSE;

    FB_TN_SC_AREA_RESTORE.Xus_TN_SCREEN := Xus_TN_SCREEN;
    FB_TN_SC_AREA_RESTORE();
    Xus_TN_SCREEN := FB_TN_SC_AREA_RESTORE.Xus_TN_SCREEN;

    Xus_TN_SCREEN.bo_Modal_Dialog := FALSE;
  END_IF;

END_FUNCTION_BLOCK

(* ---- 720-HEAT_METER.ST ---- *)
FUNCTION UDINT_TO_TIME2:TIME
	VAR_INPUT
		IN :	UDINT;
	END_VAR
	UDINT_TO_TIME2 := DINT_TO_TIME(UDINT_TO_DINT(IN));
END_FUNCTION

FUNCTION_BLOCK T_PLC_MS_block
	VAR_OUTPUT
		T_PLC_MS :	UDINT;
	END_VAR

	VAR_EXTERNAL
		PLC_TICKS_PER_SEC :	INT;
		PLC_SYS_TICK_CNT :	DINT;
	END_VAR

	VAR
		debug :	BOOL;(*Debug-Mode ON / OFF*)
		N :	INT;(*Debug-Faktor*)
		Offset :	UDINT;(*Debug-Offset*)
		temp :	DWORD := DWORD#1;(*Debug-Offset*)
		mode :	BOOL;(*modus*)
		faktor :	UDINT;(*Systemtakt-Faktor*)
		init :	BOOL;
		v_plc_ticks_per_sec :	UDINT;
		base :	UDINT := UDINT#1000;
	END_VAR

	IF init = FALSE THEN
		v_plc_ticks_per_sec := INT_TO_UDINT(PLC_TICKS_PER_SEC);
		IF v_plc_ticks_per_sec = UDINT#1024 THEN
			faktor := UDINT#1;
			mode := FALSE;
		ELSIF v_plc_ticks_per_sec > UDINT#0 THEN
			IF v_plc_ticks_per_sec <= base THEN
				faktor := base / v_plc_ticks_per_sec;
				mode := FALSE;
			ELSE
				faktor := v_plc_ticks_per_sec / base;
				mode := TRUE;
			END_IF;
		ELSE
			faktor := UDINT#1;
		END_IF;
		init := TRUE;
	END_IF;

	IF mode THEN
		T_PLC_MS := DINT_TO_UDINT(PLC_SYS_TICK_CNT) / faktor;
	ELSE
		T_PLC_MS := DINT_TO_UDINT(PLC_SYS_TICK_CNT) * faktor;
	END_IF;

	IF debug THEN
		T_PLC_MS := (DWORD_TO_UDINT(SHL(UDINT_TO_DWORD(T_PLC_MS),N) OR SHL(temp,N)) - UDINT#1) + Offset;
	END_IF;

END_FUNCTION_BLOCK

TYPE
	oscat_ARRAY_X               : ARRAY [0..1]    OF REAL;
	oscat_XY                    : ARRAY [1..20]   OF oscat_ARRAY_X := [0,0,0,0,0,0,0,0,0,0,0,0,0,0,0,0,0,0,0,0];
END_TYPE

FUNCTION_BLOCK LINEAR_INT_Block

	VAR_INPUT
		X :	REAL;
		XY :	oscat_XY;
		PTS :	INT;
	END_VAR

	VAR_OUTPUT
		LINEAR_INT :	REAL;
	END_VAR

	VAR
		i :	INT;
		i2 :	INT;
	END_VAR

	pts := MIN(pts,20);

	i := 2;

	WHILE (i < pts) AND (XY[i][0] < X) DO
		i := i + 1;
	END_WHILE;

	i2 := i-1;

	LINEAR_INT := ((XY[i][1] - XY[i2][1]) * X - XY[i][1] * XY[i2][0] + XY[i2][1] * XY[i][0]) / (XY[i][0] - XY[i2][0]);

END_FUNCTION_BLOCK

FUNCTION_BLOCK WATER_ENTHALPY_Block

    VAR_INPUT
        T :	REAL;
    END_VAR

    VAR_OUTPUT
        RESULT :	REAL;
    END_VAR

    VAR
        Pts :	INT;
        data :	oscat_XY;
        FB_LINEAR_INT :	LINEAR_INT_Block;
    END_VAR

    IF Pts = 0 THEN
        Pts := 11;
        data[01][0] := REAL#0.0;
        data[01][1] := REAL#0.06;
        data[02][0] := REAL#10.0;
        data[02][1] := REAL#42.1;
        data[03][0] := REAL#20.0;
        data[03][1] := REAL#83.9;
        data[04][0] := REAL#30.0;
        data[04][1] := REAL#125.8;
        data[05][0] := REAL#40.0;
        data[05][1] := REAL#167.58;
        data[06][0] := REAL#50.0;
        data[06][1] := REAL#209.4;
        data[07][0] := REAL#60.0;
        data[07][1] := REAL#251.2;
        data[08][0] := REAL#70.0;
        data[08][1] := REAL#293.1;
        data[09][0] := REAL#80.0;
        data[09][1] := REAL#335.0;
        data[10][0] := REAL#90.0;
        data[10][1] := REAL#377.0;
        data[11][0] := REAL#100.0;
        data[11][1] := REAL#419.1;
    END_IF;

    FB_LINEAR_INT(X:=T,XY:=Data,Pts:=Pts);
    Result :=FB_LINEAR_INT.LINEAR_INT;

END_FUNCTION_BLOCK

FUNCTION_BLOCK R2_SET_Block

	VAR_INPUT
		X :	REAL;
	END_VAR

	VAR_OUTPUT
		R2_SET :	REAL2;
	END_VAR

	R2_SET.RX := X;
	R2_SET.R1 := 0.0;

END_FUNCTION_BLOCK

FUNCTION_BLOCK R2_ADD_Block

	VAR_INPUT
		X :	REAL2;
		Y :	REAL;
	END_VAR

	VAR_OUTPUT
		R2_ADD :	REAL2;
	END_VAR

	VAR
		temp :	REAL;
	END_VAR

	temp := X.RX;
	R2_ADD.RX := Y + X.R1 + X.RX;
	R2_ADD.R1 := temp - R2_ADD.RX + Y + X.R1;

END_FUNCTION_BLOCK

TYPE REAL2:

	STRUCT
		R1 : REAL;
		RX : REAL;
	END_STRUCT;

END_TYPE

FUNCTION_BLOCK INTEGRATE

	VAR_INPUT
		E :	BOOL := TRUE;
		X :	REAL;
		K :	REAL := 1.0;
	END_VAR

	VAR_IN_OUT
		Y :	REAL;
	END_VAR

	VAR
		X_last :	REAL;
		init :	BOOL;
		T_PLC_MS :	T_PLC_MS_block;
		last :	UDINT;
		tx :	UDINT;
	END_VAR

	T_PLC_MS();
	tx:= T_PLC_MS.T_PLC_MS;

	IF NOT init THEN
		init := TRUE;
		X_last := X;
	ELSIF E THEN
		Y := (X + X_LAST) * 0.5E-3 * UDINT_TO_REAL(tx-last) * K + Y;
		X_last := X;
	END_IF;
	last := tx;

END_FUNCTION_BLOCK

FUNCTION_BLOCK FT_INT2_Block

	VAR_INPUT
		IN :	REAL;
		K :	REAL := 1.0;
		RUN :	BOOL := TRUE;
		RST :	BOOL;
		OUT_MIN :	REAL := REAL#-1.0E-37;
		OUT_MAX :	REAL := REAL#1.0E37;
	END_VAR

	VAR_OUTPUT
		OUT :	REAL;
		LIM :	BOOL;
	END_VAR

	VAR
		integ :	INTEGRATE;
		ix :	REAL;
		val :	REAL2;
		R2_ADD :	R2_ADD_Block;
		R2_SET :	R2_SET_Block;
	END_VAR

	IF RST THEN
		R2_SET(X:=0.0);
		val:=R2_SET.R2_SET;
		out := 0.0;
	ELSE
		integ(X := IN, E := RUN, K := K, Y := ix);
		ix := integ.Y;
		R2_ADD(X:=val,Y:=ix);
		val:=R2_ADD.R2_ADD;
		ix := 0.0;
		OUT := val.RX;
	END_IF;

	(* check output for limits *)
	IF out > OUT_MIN AND out < OUT_MAX THEN
		LIM := FALSE;
	ELSE
		OUT := LIMIT(OUT_MIN, OUT, OUT_MAX);
		R2_SET(X:=OUT);
		val:=R2_SET.R2_SET;
		LIM := TRUE;
	END_IF;

END_FUNCTION_BLOCK

FUNCTION WATER_DENSITY:REAL

    VAR_INPUT
        T :	REAL;
        SAT :	BOOL;
    END_VAR

    VAR
        T2 :	REAL;
        T4 :	REAL;
    END_VAR

    T2 := T * T;
    T4 := T2 * T2;
    WATER_DENSITY := (999.83952 + 16.952577*T + -7.9905127E-3*T2 + -4.6241757E-5*T2*T + 1.0584601E-7*T4 + -2.8103006E-10*T4*T) / (1.0 + 0.0168872*T);
    IF sat THEN WATER_DENSITY := WATER_DENSITY - 0.004612 + 0.000106 * T; END_IF;

END_FUNCTION

FUNCTION TIME_TO_UDINT2:UDINT
	VAR_INPUT
		X :	TIME;
	END_VAR

	TIME_TO_UDINT2 := DINT_TO_UDINT(TIME_TO_DINT(X));
END_FUNCTION

FUNCTION_BLOCK HEAT_METER_Block

	VAR_INPUT
		TF :	REAL;
		TR :	REAL;
		LPH :	REAL;
		E :	BOOL;
		RST :	BOOL;
		CP :	REAL;
		DENSITY :	REAL;
		CONTENT :	REAL;
		PULSE_MODE :	BOOL;
		RETURN_METER :	BOOL;
		AVG_TIME :	TIME := T#5s;
	END_VAR

	VAR_OUTPUT
		C :	REAL;
	END_VAR

	VAR_IN_OUT
		Y :	REAL;
	END_VAR

	VAR
		tx :	UDINT;
		last :	UDINT;
		int1 :	FT_INT2_Block;
		edge :	BOOL;
		x :	REAL;
		init :	BOOL;
		Y_last :	REAL;
		T_PLC_MS :	T_PLC_MS_Block;
		WATER_ENTHALPY :	WATER_ENTHALPY_Block;
		wa_TF :	REAL;
		wa_TR :	REAL;
	END_VAR

	IF rst THEN
		int1(rst := TRUE);
		int1.rst := FALSE;
		C := 0.0;
		Y := 0.0;
	ELSIF e THEN
		water_enthalpy(T:=TF);
		wa_TF:=water_enthalpy.Result;

		water_enthalpy(T:=TR);
		wa_TR:=water_enthalpy.Result;

		X := (WATER_DENSITY(SEL(return_meter, TF, TR), FALSE) * (wa_TF - wa_TR) * (1.0 - content) + CP * Density * content * (TF-TR));
	END_IF;

	int1(run := NOT pulse_mode AND e, in := X * LPH * 2.77777777777E-4);
	IF pulse_mode THEN
		IF NOT edge AND E THEN Y := Y + X * LPH; END_IF;
	ELSE
		Y := int1.Out;
	END_IF;

	edge := e;

	T_PLC_MS();
	tx:= T_PLC_MS.T_PLC_MS;

	IF NOT init THEN
		init := TRUE;
		last := tx;
	END_IF;

	IF (tx - last >= TIME_TO_UDINT2(AVG_TIME)) AND (avg_time > T#0s) THEN
		last := tx;
		C := (Y - Y_last) * 3.6E12 / TIME_TO_REAL(AVG_TIME);
		Y_last := Y;
	END_IF;

END_FUNCTION_BLOCK

PROGRAM program0
	VAR
	    TF :	REAL;
		TR :	REAL;
		LPH :	REAL;
		E :	BOOL;
		RST :	BOOL;
		CP :	REAL;
		DENSITY :	REAL;
		CONTENT :	REAL;
		PULSE_MODE :	BOOL;
		RETURN_METER :	BOOL;
		AVG_TIME :	TIME := T#5s;
		Y :	REAL;
		C :	REAL;

		func_block : HEAT_METER_Block;
  	END_VAR
	func_block.TF := TF;
	func_block.TR := TR;
	func_block.LPH := LPH;
	func_block.E := E;
	func_block.RST := RST;
	func_block.CP := CP;
	func_block.DENSITY := DENSITY;
	func_block.CONTENT := CONTENT;
	func_block.PULSE_MODE := PULSE_MODE;
	func_block.RETURN_METER := RETURN_METER;
	func_block.AVG_TIME := AVG_TIME;
	func_block.Y := Y;

	func_block();
	Y := func_block.Y;
	C := func_block.C;
END_PROGRAM

CONFIGURATION Config0
	VAR_GLOBAL
		PLC_TICKS_PER_SEC :	INT;
		PLC_SYS_TICK_CNT :	DINT;
	END_VAR
  	RESOURCE Res0 ON PLC
    	TASK task0(INTERVAL := T#20ms,PRIORITY := 0);
    	PROGRAM instance0 WITH task0 : program0;
  	END_RESOURCE
END_CONFIGURATION

(* ---- 721-FILE_SERVER.ST ---- *)
FUNCTION_BLOCK FILE_SERVER_Block

	VAR
		buf_size :	UDINT := UDINT#4096;
		handle :	UINT;
		read_max_length :	UDINT;
		file_position :	UDINT;
		used_filename :	STRING;
		close_time :	TIME;
		length_read :	UDINT;
		write_length :	UDINT;
		length_written :	UDINT;
		open_handle :	UINT;
		seek_mode :	UINT;
		seek_position :	UDINT;
		tell_position :	UDINT;
	END_VAR

	VAR
		last_mode :	BYTE;
		command :	BYTE;
		error_code :	BYTE;
		error :	BOOL;
		file_change :	BOOL;
		step :	INT;
		t_diff :	TIME;
		tx_last :	TIME;
		tx :	TIME;
	END_VAR

	VAR_IN_OUT
		FSD :	oscat_FILE_SERVER_DATA;
		PT :	oscat_NETWORK_BUFFER;
	END_VAR

	VAR
		FILE_REMOVE :	FILE_REMOVE;
		FILE_OPEN :	FILE_OPEN;
		FILE_SEEK :	FILE_SEEK;
		FILE_TELL :	FILE_TELL;
		FILE_CLOSE :	FILE_CLOSE;
		FILE_READ :	FILE_READ;
		FILE_WRITE :	FILE_WRITE;
		T_PLC_MS :	T_PLC_MS;
	END_VAR

	T_PLC_MS();
	tx := UDINT_TO_TIME(T_PLC_MS.T_PLC_MS);
	t_diff := tx - tx_last;
	tx_last := tx;

	CASE step OF
	0:
		IF FSD.MODE = LIMIT(BYTE#1,FSD.MODE,BYTE#5) THEN
			close_time := T#1ms;
			IF handle = UINT#00 AND FSD.MODE <= BYTE#3 THEN
				step := 100;
			ELSE
				IF EQ_STRING(used_filename, FSD.FILENAME) AND FSD.MODE = last_mode THEN
					step := 200;
				ELSE
					step := 32000;
					file_change := FSD.MODE <> BYTE#5;
				END_IF;
			END_IF;
		ELSIF handle > UINT#0 THEN
			IF FSD.AUTO_CLOSE > T#0s THEN
				close_time := close_time + t_diff;
				IF close_time > FSD.AUTO_CLOSE THEN
					step := 32000;
				END_IF;
			END_IF;
		END_IF;

	100:
		IF FSD.MODE = BYTE#3 OR FSD.MODE = BYTE#4 THEN
			command := BYTE#7;
			step := 110;
		ELSE
			step := 120;
		END_IF;

	110:
		IF command = BYTE#0  THEN
			IF (FSD.MODE = BYTE#4) OR (error and error_code <> BYTE#143) THEN
				step := 30000;
			ELSE
				step := 120;
			END_IF;
		END_IF;

	120:
		command := BYTE#1;
		last_mode := FSD.MODE;
		step := 122;

	122:
		IF command = BYTE#0 THEN
			IF error THEN
				step := 30000;
			ELSE

				close_time := T#1ms;
				handle := open_handle;
				used_filename := FSD.FILENAME;
				file_position := UDINT#4294967295;
				FSD.FILE_SIZE := UDINT#0;
				step := 125;
			END_IF;
		END_IF;

	125:
		seek_mode := UINT#2;
		seek_position := UDINT#0;
		command := BYTE#5;
		step := 130;

	130:
		IF command = BYTE#0 THEN
			IF Error THEN
				step := 30000;
			ELSE
				step := 140;
			END_IF;
		END_IF;

	140:
		command := BYTE#6;
		step := 150;

	150:
		IF command = BYTE#0 THEN
			IF Error THEN
				step := 30000;
			ELSE
				FSD.FILE_SIZE := tell_position;
				file_position := tell_position;
				FSD.FILE_OPEN := TRUE;
				step := 200;
			END_IF;
		END_IF;

	200:
		IF FSD.OFFSET > FSD.FILE_SIZE THEN
			error_code := BYTE#255;
			step := 30000;
		ELSIF FSD.OFFSET <> file_position THEN
			command := BYTE#5;
			seek_mode := UINT#0;
			seek_position := FSD.OFFSET;
			step := 210;
		ELSE
			step := 300;
		END_IF;

	210:
		IF command = BYTE#0 THEN
			file_position := seek_position;
			IF Error THEN
				step := 30000;
			ELSE
				step := 300;
			END_IF;
		END_IF;

	300:
		IF FSD.MODE = BYTE#1 THEN
			step := 400;
		ELSE
			step := 500;
		END_IF;

	400:
		IF UINT_TO_UDINT(PT.SIZE) > buf_size THEN
			read_max_length := buf_size;
		ELSE
			read_max_length := UINT_TO_UDINT(PT.SIZE);
		END_IF;

		IF file_position + read_max_length > FSD.FILE_SIZE THEN
			read_max_length := FSD.FILE_SIZE - file_position;
		END_IF;

		IF read_max_length > UDINT#0 THEN
			command := BYTE#3;
			step := INT#410;
		ELSE
			PT.SIZE := UINT#0;
			step := 30000;
		END_IF;

	410:
		IF command = BYTE#0 THEN
			PT.SIZE := UDINT_TO_UINT(length_read);
			IF NOT Error THEN
				file_position := file_position + length_read;
				FSD.OFFSET := file_position;
			END_IF;
			step := 30000;
		END_IF;

	500:
		IF UINT_TO_UDINT(PT.SIZE) > buf_size THEN
			write_length := buf_size;
		ELSE
			write_length := UINT_TO_UDINT(PT.SIZE);
		END_IF;

		IF write_length > UDINT#0 THEN
			command := BYTE#4;
			step := INT#510;
		ELSE
			step := 30000;
		END_IF;

	510:
		IF command = BYTE#0 THEN
			IF NOT Error THEN
				file_position := file_position + length_written;
				FSD.OFFSET := file_position;
				IF file_position > FSD.FILE_SIZE THEN
					FSD.FILE_SIZE := file_position;
				END_IF;
			END_IF;
			step := 30000;
		END_IF;

	30000:
		FSD.MODE := BYTE#0;
		FSD.ERROR := error_code;
		step := 0;

	32000:
		close_time := T#0s;
		IF handle > UINT#0 THEN
			command := BYTE#2;
		END_IF;
		step := 32100;

	32100:
		IF command = BYTE#0 THEN
			FSD.FILE_OPEN := FALSE;
			file_position := UDINT#0;
			FSD.FILE_SIZE := UDINT#0;
			FSD.OFFSET := UDINT#0;
			used_filename := '';
			handle := UINT#00;

			IF file_change THEN
				file_change := FALSE;
				step := 100;
			ELSE
				step := 30000;
			END_IF;
		END_IF;

	END_CASE;

	FILE_OPEN.Execute := command = BYTE#1;
	FILE_OPEN.Name := FSD.FILENAME;
	FILE_OPEN();
	open_handle := FILE_OPEN.Handle;

	IF command = BYTE#1 THEN
		IF FILE_OPEN.Done THEN
			error := FILE_OPEN.Error;
			command := BYTE#0;
			error_code := SEL_BYTE(error,BYTE#00,UINT_TO_BYTE(FILE_OPEN.ErrorID));
		END_IF;
	END_IF;

	FILE_CLOSE.Execute := command = BYTE#2;
	FILE_CLOSE.Handle := Handle;
	FILE_CLOSE();

	IF command = BYTE#2 THEN
		IF FILE_CLOSE.Done THEN
			error := FILE_CLOSE.Error;
			command := BYTE#0;
			error_code := SEL_BYTE(error,BYTE#00,UINT_TO_BYTE(FILE_CLOSE.ErrorID + UINT#10));
		END_IF;
	END_IF;

	FILE_READ.Execute := command = BYTE#3;
	FILE_READ.Handle := handle;
	FILE_READ.MaxLength := read_max_length;
	FILE_READ.Buffer := PT.BUFFER;
	FILE_READ();
	PT.BUFFER := FILE_READ.Buffer;

	IF command = BYTE#3 THEN
		IF FILE_READ.Done THEN
			error := FILE_READ.Error;
			command := BYTE#0;
			length_read :=  FILE_READ.LengthRead;
			error_code := SEL_BYTE(error,BYTE#00,UINT_TO_BYTE(FILE_READ.ErrorID + UINT#40));
		END_IF;
	END_IF;

	FILE_WRITE.Execute   := command = BYTE#4;
	FILE_WRITE.Handle    := handle;
	FILE_WRITE.Length    := write_length ;
	FILE_WRITE.Buffer    := PT.BUFFER;
	FILE_WRITE();
	PT.BUFFER := FILE_WRITE.Buffer;

	IF command = BYTE#4 THEN
		IF FILE_WRITE.Done THEN
			error := FILE_WRITE.Error;
			command := BYTE#0;
			length_written := write_length;
			error_code := SEL_BYTE(error,BYTE#00,UINT_TO_BYTE(FILE_WRITE.ErrorID + UINT#70));
		END_IF;
	END_IF;

	FILE_SEEK.Execute  := command = BYTE#5;
	FILE_SEEK.Handle   := handle;
	FILE_SEEK.Mode     := seek_mode;
	FILE_SEEK.Position := UDINT_TO_DINT(seek_position);
	FILE_SEEK();

	IF command = BYTE#5 THEN
		IF FILE_SEEK.Done THEN
			error := FILE_SEEK.Error;
			command := BYTE#0;
			error_code := SEL_BYTE(error,BYTE#00,UINT_TO_BYTE(FILE_SEEK.ErrorID + UINT#100));
		END_IF;
	END_IF;

	FILE_TELL.Execute := command = BYTE#6;
	FILE_TELL.Handle := handle;
	FILE_TELL();

	IF command = BYTE#6 THEN
		IF FILE_TELL.Done THEN
			error := FILE_TELL.Error;
			command := BYTE#0;
			tell_position := DINT_TO_UDINT(FILE_TELL.Position);
			error_code := SEL_BYTE(error,BYTE#00,UINT_TO_BYTE(FILE_TELL.ErrorID + UINT#130));
		END_IF;
	END_IF;

	FILE_REMOVE.Execute := command = BYTE#7;
	FILE_REMOVE.Name := FSD.FILENAME;
	FILE_REMOVE();

	IF command = BYTE#7 THEN
		IF FILE_REMOVE.Done THEN
			error := FILE_REMOVE.Error;
			command := BYTE#0;
			error_code := SEL_BYTE(error,BYTE#00,UINT_TO_BYTE(FILE_REMOVE.ErrorID + UINT#140));
		END_IF;
	END_IF;

END_FUNCTION_BLOCK

PROGRAM program0
	VAR
		FSD :	oscat_FILE_SERVER_DATA;
		PT :	oscat_NETWORK_BUFFER;

		func_block : FILE_SERVER_Block;
	END_VAR
	func_block.FSD := FSD;
	func_block.PT := PT;

	func_block();
	FSD  := func_block.FSD;
	PT  := func_block.PT;
END_PROGRAM

CONFIGURATION Config0
	RESOURCE Res0 ON PLC
		TASK task0(INTERVAL := T#20ms,PRIORITY := 0);
		PROGRAM instance0 WITH task0 : program0;
	END_RESOURCE
END_CONFIGURATION

(* ---- 722-BLIND_CONTROL_S.ST ---- *)
FUNCTION UDINT_TO_TIME2:TIME

	VAR_INPUT
		IN :	UDINT;
	END_VAR

	UDINT_TO_TIME2 := DINT_TO_TIME(UDINT_TO_DINT(IN));

END_FUNCTION

FUNCTION_BLOCK T_PLC_MS_block
	VAR_OUTPUT
		T_PLC_MS :	UDINT;
	END_VAR

	VAR_EXTERNAL
		PLC_TICKS_PER_SEC :	INT;
		PLC_SYS_TICK_CNT :	DINT;
	END_VAR

	VAR
		debug :	BOOL;(*Debug-Mode ON / OFF*)
		N :	INT;(*Debug-Faktor*)
		Offset :	UDINT;(*Debug-Offset*)
		temp :	DWORD := DWORD#1;(*Debug-Offset*)
		mode :	BOOL;(*modus*)
		faktor :	UDINT;(*Systemtakt-Faktor*)
		init :	BOOL;
		v_plc_ticks_per_sec :	UDINT;
		base :	UDINT := UDINT#1000;
	END_VAR

	IF init = FALSE THEN
		v_plc_ticks_per_sec := INT_TO_UDINT(PLC_TICKS_PER_SEC);
		IF v_plc_ticks_per_sec = UDINT#1024 THEN
			faktor := UDINT#1;
			mode := FALSE;
		ELSIF v_plc_ticks_per_sec > UDINT#0 THEN
			IF v_plc_ticks_per_sec <= base THEN
				faktor := base / v_plc_ticks_per_sec;
				mode := FALSE;
			ELSE
				faktor := v_plc_ticks_per_sec / base;
				mode := TRUE;
			END_IF;
		ELSE
			faktor := UDINT#1;
		END_IF;
		init := TRUE;
	END_IF;

	IF mode THEN
		T_PLC_MS := DINT_TO_UDINT(PLC_SYS_TICK_CNT) / faktor;
	ELSE
		T_PLC_MS := DINT_TO_UDINT(PLC_SYS_TICK_CNT) * faktor;
	END_IF;

	IF debug THEN
		T_PLC_MS := (DWORD_TO_UDINT(SHL(UDINT_TO_DWORD(T_PLC_MS),N) OR SHL(temp,N)) - UDINT#1) + Offset;
	END_IF;
END_FUNCTION_BLOCK

FUNCTION TIME_TO_UDINT2:UDINT
	VAR_INPUT
		X :	TIME;
	END_VAR

	TIME_TO_UDINT2 := DINT_TO_UDINT(TIME_TO_DINT(X));
END_FUNCTION

FUNCTION FRMP_B:BYTE
	VAR_INPUT
		START :	BYTE;
		DIR :	BOOL;
		TD :	TIME;
		TR :	TIME;
	END_VAR

	IF TD < TR THEN
		FRMP_B := MIN(UDINT_TO_BYTE(DWORD_TO_UDINT(SHL(TIME_TO_DWORD(TD), 8)) / TIME_TO_UDINT2(TR)), SEL(DIR, START, USINT_TO_BYTE(USINT#255 - BYTE_TO_USINT(START))));
		IF DIR THEN
			FRMP_B := USINT_TO_BYTE(BYTE_TO_USINT(START) + BYTE_TO_USINT(FRMP_B));
		ELSE
			FRMP_B := USINT_TO_BYTE(BYTE_TO_USINT(START) - BYTE_TO_USINT(FRMP_B));
		END_IF;
	ELSE
		FRMP_B := SEL(DIR, BYTE#0, BYTE#255);
	END_IF;
END_FUNCTION

FUNCTION_BLOCK _RMP_B
	VAR_INPUT
		DIR :	BOOL;
		E :	BOOL := TRUE;
		TR :	TIME;
	END_VAR

	VAR_IN_OUT
		RMP :	BYTE;
	END_VAR

	VAR
		T_PLC_MS :	T_PLC_MS_block;
		tx :	TIME;
		tl :	TIME;
		tn :	TIME;
		init :	BOOL;
		last_dir :	BOOL;
		start :	BYTE;
	END_VAR

	T_PLC_MS();
	tx := UDINT_TO_TIME(T_PLC_MS.T_PLC_MS);

	IF E AND init AND (dir = last_dir) AND (RMP <> SEL(DIR, BYTE#0, BYTE#255)) AND TR = tn THEN
		RMP := FRMP_B(start, DIR, tx - tl, TR);
	ELSE
		init := TRUE;
		tl := tx;
		tn := tr;
		start := RMP;
	END_IF;
	last_dir := dir;
END_FUNCTION_BLOCK

FUNCTION_BLOCK TREND_DW
	VAR_INPUT
		X :	DWORD;
	END_VAR
	VAR_OUTPUT
		Q :	BOOL;
		TU :	BOOL;
		TD :	BOOL;
		D :	DWORD;
	END_VAR

	VAR
		LAST_X :	DWORD;
	END_VAR

	IF X > last_X THEN
		TU := TRUE;
		TD := FALSE;
		D := UDINT_TO_DWORD(DWORD_TO_UDINT(X) - DWORD_TO_UDINT(last_X));
		Q := TRUE;
	ELSIF X < last_X THEN
		TD := TRUE;
		TU := FALSE;
		D := UDINT_TO_DWORD(DWORD_TO_UDINT(last_X) - DWORD_TO_UDINT(X));
		Q := FALSE;
	ELSE
		TU := FALSE;
		TD := FALSE;
		D := DWORD#0;
	END_IF;
	last_X := X;
END_FUNCTION_BLOCK

FUNCTION_BLOCK _RMP_NEXT
	VAR_INPUT
		E :	BOOL := TRUE;
		IN :	BYTE;
		TR :	TIME;
		TF :	TIME;
		TL :	TIME;
	END_VAR

	VAR_OUTPUT
		DIR :	BOOL;
		UP :	BOOL;
		DN :	BOOL;
	END_VAR

	VAR_IN_OUT
		OUT :	BYTE;
	END_VAR
	VAR
		rmx :	_RMP_B;
		dirx :	TREND_DW;
		t_lock :	TP;
		xen :	BOOL;
		xdir :	BOOL;
	END_VAR

	dirx(X := BYTE_TO_DWORD(in));

	t_lock(in := FALSE, pt := TL);

	IF dirx.TU AND (OUT < IN) THEN
		IF NOT xdir AND xen THEN t_lock(in := TRUE); END_IF;
		xen := TRUE;
		xdir := TRUE;
	ELSIF dirx.TD AND (OUT > IN) THEN
		IF xdir AND xen THEN t_lock(in := TRUE); END_IF;
		xen := TRUE;
		xdir := FALSE;
	ELSIF xen THEN
		IF (xdir AND (out >= in)) OR (NOT xdir AND (out <= in)) THEN
			xen := FALSE;
			IF tl > t#0s THEN t_lock(IN := TRUE); END_IF;
		END_IF;
	END_IF;

	IF NOT t_lock.Q AND xen THEN
		UP := XDIR;
		DIR := XDIR;
		DN := NOT XDIR;
	ELSE
		UP := FALSE;
		DN := FALSE;
	END_IF;

	rmx(rmp := OUT, E := E AND (UP OR DN) , dir := DIR, tr := SEL(dir, TF, TR));
	OUT := rmx.RMP;
END_FUNCTION_BLOCK

FUNCTION _BYTE_TO_INT:INT
	VAR_INPUT
		IN :	BYTE;
	END_VAR

	_BYTE_TO_INT := USINT_TO_INT(BYTE_TO_USINT(IN));
END_FUNCTION

FUNCTION_BLOCK BLIND_CONTROL_S_Block

	VAR_INPUT
		UP :	BOOL;
		DN :	BOOL;
		S_IN :	BYTE := BYTE#125;
		PI :	BYTE;
		T_UP :	TIME;
		T_DN :	TIME;
		RU :	BOOL;
		RD :	BOOL;
		T_LOCKOUT :	TIME := T#100ms;
		T_EXT :	TIME;
		EXT_TRIG :	BYTE := BYTE#5;
		R_POS_TOP :	BYTE := BYTE#255;
		R_POS_BOT :	BYTE;
	END_VAR

	VAR_OUTPUT
		POS :	BYTE;
		MU :	BOOL;
		MD :	BOOL;
		STATUS :	BYTE;
	END_VAR

	VAR
		T_PLC_MS :	T_PLC_MS_Block;
		rmp :	_RMP_NEXT;
		tx :	TIME;
		last :	TIME;
		pi_last :	BYTE;
	END_VAR

	T_PLC_MS();
	tx:= UDINT_TO_TIME(T_PLC_MS.T_PLC_MS);

	IF UP  AND NOT DN THEN
		rmp.IN := BYTE#255;
		STATUS := BYTE#121;
	ELSIF DN AND NOT UP THEN
		rmp.IN := BYTE#0;
		STATUS := BYTE#122;
	ELSIF NOT (UP OR DN) THEN
		rmp.IN := PI;
		STATUS := S_IN;
	END_IF;

	rmp(E := UP OR DN, TR := T_UP, TF := T_DN, TL := T_LOCKOUT, OUT := POS);
	pos := rmp.OUT;

	CASE _BYTE_TO_INT(STATUS) OF
		0:
			last := tx;
			PI_last := PI XOR BYTE#255;
			STATUS := BYTE#128;

		121:
			MU := TRUE;
			MD := FALSE;
			IF POS >= USINT_TO_BYTE(USINT#255 - BYTE_TO_USINT(EXT_TRIG)) THEN
				POS := BYTE#255;
				last := tx;
				STATUS := BYTE#129;
			END_IF;

		122:
			MD := TRUE;
			MU := FALSE;
			IF POS <= EXT_TRIG THEN
				POS := BYTE#0;
				last := tx;
				STATUS := BYTE#129;
			END_IF;

		123:
			MD := rmp.DN;
			MU := rmp.UP;
			IF NOT (rmp.DN OR rmp.UP) THEN
				IF POS <= EXT_TRIG THEN
					MD := TRUE;
					last := tx;
					STATUS := BYTE#129;
				ELSIF POS >= USINT_TO_BYTE(USINT#255 - BYTE_TO_USINT(EXT_TRIG)) THEN
					MU := TRUE;
					last := tx;
					STATUS := BYTE#129;
				ELSE
					STATUS := S_IN;
				END_IF;
			END_IF;

		124:
			MD := rmp.DN;
			MU := rmp.UP;
			IF NOT(rmp.DN OR rmp.UP) THEN
				PI_last := PI;
				STATUS := S_IN;
			END_IF;

		127:
			IF (tx - last) >= T_LOCKOUT THEN
					STATUS := S_IN;
			END_IF;

		128:
			MU := TRUE;
			MD := FALSE;
			rmp.IN := BYTE#255;
			IF (tx - last) >= (T_UP +  T_EXT) THEN
				MU := FALSE;
				last := tx;
				STATUS := BYTE#127;
			END_IF;

		129:
			IF (tx - last) >= T_EXT THEN
				MU := FALSE;
				MD := FALSE;
				last := tx;
				STATUS := BYTE#127;
			END_IF;

	ELSE
		MU := FALSE;
		MD := FALSE;
		IF PI <> PI_last THEN
			PI_last := PI;
			rmp.IN := PI;
			STATUS := BYTE#123;
		ELSIF POS = BYTE#0 AND RU THEN
			rmp.IN := R_POS_BOT;
			STATUS := BYTE#124;
		ELSIF pos = BYTE#255 AND RD THEN
			rmp.IN := R_POS_TOP;
			STATUS := BYTE#124;
		ELSE
			STATUS := S_IN;
		END_IF;
	END_CASE;

END_FUNCTION_BLOCK

PROGRAM program0
	VAR
		UP :	BOOL;
		DN :	BOOL;
		S_IN :	BYTE := BYTE#125;
		PI :	BYTE;
		T_UP :	TIME;
		T_DN :	TIME;
		RU :	BOOL;
		RD :	BOOL;
		T_LOCKOUT :	TIME := T#100ms;
		T_EXT :	TIME;
		EXT_TRIG :	BYTE := BYTE#5;
		R_POS_TOP :	BYTE := BYTE#255;
		R_POS_BOT :	BYTE;
		POS :	BYTE;
		MU :	BOOL;
		MD :	BOOL;
		STATUS :	BYTE;
		func_block : BLIND_CONTROL_S_Block;
	END_VAR
	func_block.UP := UP;
	func_block.DN := DN;
	func_block.S_IN := S_IN ;
	func_block.PI    := PI    ;
	func_block.T_UP := T_UP;
	func_block.T_DN := T_DN ;
	func_block.RU    := RU    ;
	func_block.RD := RD;
	func_block.T_LOCKOUT := T_LOCKOUT;
	func_block.T_EXT := T_EXT ;
	func_block.EXT_TRIG    := EXT_TRIG    ;
	func_block.R_POS_TOP := R_POS_TOP;
	func_block.R_POS_BOT := R_POS_BOT ;
	func_block();
	POS  := func_block.POS;
	MU  := func_block.MU;
	MD  := func_block.MD;
	STATUS  := func_block.STATUS;
END_PROGRAM

CONFIGURATION Config0
	VAR_GLOBAL
		PLC_TICKS_PER_SEC :	INT;
		PLC_SYS_TICK_CNT :	DINT;
	END_VAR
  	RESOURCE Res0 ON PLC
    	TASK task0(INTERVAL := T#20ms,PRIORITY := 0);
    	PROGRAM instance0 WITH task0 : program0;
  	END_RESOURCE
END_CONFIGURATION

(* ---- 723-ACTUATOR_3P.ST ---- *)
FUNCTION UDINT_TO_TIME2:TIME

	VAR_INPUT
		IN :	UDINT;
	END_VAR

	UDINT_TO_TIME2 := DINT_TO_TIME(UDINT_TO_DINT(IN));

END_FUNCTION

FUNCTION_BLOCK T_PLC_MS_block
	VAR_OUTPUT
		T_PLC_MS :	UDINT;
	END_VAR

	VAR_EXTERNAL
		PLC_TICKS_PER_SEC :	INT;
		PLC_SYS_TICK_CNT :	DINT;
	END_VAR

	VAR
		debug :	BOOL;(*Debug-Mode ON / OFF*)
		N :	INT;(*Debug-Faktor*)
		Offset :	UDINT;(*Debug-Offset*)
		temp :	DWORD := DWORD#1;(*Debug-Offset*)
		mode :	BOOL;(*modus*)
		faktor :	UDINT;(*Systemtakt-Faktor*)
		init :	BOOL;
		v_plc_ticks_per_sec :	UDINT;
		base :	UDINT := UDINT#1000;
	END_VAR

	IF init = FALSE THEN
		v_plc_ticks_per_sec := INT_TO_UDINT(PLC_TICKS_PER_SEC);
		IF v_plc_ticks_per_sec = UDINT#1024 THEN
			faktor := UDINT#1;
			mode := FALSE;
		ELSIF v_plc_ticks_per_sec > UDINT#0 THEN
			IF v_plc_ticks_per_sec <= base THEN
				faktor := base / v_plc_ticks_per_sec;
				mode := FALSE;
			ELSE
				faktor := v_plc_ticks_per_sec / base;
				mode := TRUE;
			END_IF;
		ELSE
			faktor := UDINT#1;
		END_IF;
		init := TRUE;
	END_IF;

	IF mode THEN
		T_PLC_MS := DINT_TO_UDINT(PLC_SYS_TICK_CNT) / faktor;
	ELSE
		T_PLC_MS := DINT_TO_UDINT(PLC_SYS_TICK_CNT) * faktor;
	END_IF;

	IF debug THEN
		T_PLC_MS := (DWORD_TO_UDINT(SHL(UDINT_TO_DWORD(T_PLC_MS),N) OR SHL(temp,N)) - UDINT#1) + Offset;
	END_IF;
END_FUNCTION_BLOCK

FUNCTION TIME_TO_UDINT2:UDINT
	VAR_INPUT
		X :	TIME;
	END_VAR

	TIME_TO_UDINT2 := DINT_TO_UDINT(TIME_TO_DINT(X));
END_FUNCTION

FUNCTION FRMP_B:BYTE
	VAR_INPUT
		START :	BYTE;
		DIR :	BOOL;
		TD :	TIME;
		TR :	TIME;
	END_VAR

	IF TD < TR THEN
		FRMP_B := MIN(UDINT_TO_BYTE(DWORD_TO_UDINT(SHL(TIME_TO_DWORD(TD), 8)) / TIME_TO_UDINT2(TR)), SEL(DIR, START, USINT_TO_BYTE(USINT#255 - BYTE_TO_USINT(START))));
		IF DIR THEN
			FRMP_B := USINT_TO_BYTE(BYTE_TO_USINT(START) + BYTE_TO_USINT(FRMP_B));
		ELSE
			FRMP_B := USINT_TO_BYTE(BYTE_TO_USINT(START) - BYTE_TO_USINT(FRMP_B));
		END_IF;
	ELSE
		FRMP_B := SEL(DIR, BYTE#0, BYTE#255);
	END_IF;
END_FUNCTION

FUNCTION_BLOCK _RMP_B
	VAR_INPUT
		DIR :	BOOL;
		E :	BOOL := TRUE;
		TR :	TIME;
	END_VAR

	VAR_IN_OUT
		RMP :	BYTE;
	END_VAR

	VAR
		T_PLC_MS :	T_PLC_MS_block;
		tx :	TIME;
		tl :	TIME;
		tn :	TIME;
		init :	BOOL;
		last_dir :	BOOL;
		start :	BYTE;
	END_VAR

	T_PLC_MS();
	tx := UDINT_TO_TIME(T_PLC_MS.T_PLC_MS);

	IF E AND init AND (dir = last_dir) AND (RMP <> SEL(DIR, BYTE#0, BYTE#255)) AND TR = tn THEN
		RMP := FRMP_B(start, DIR, tx - tl, TR);
	ELSE
		init := TRUE;
		tl := tx;
		tn := tr;
		start := RMP;
	END_IF;
	last_dir := dir;
END_FUNCTION_BLOCK

FUNCTION_BLOCK TREND_DW
	VAR_INPUT
		X :	DWORD;
	END_VAR
	VAR_OUTPUT
		Q :	BOOL;
		TU :	BOOL;
		TD :	BOOL;
		D :	DWORD;
	END_VAR

	VAR
		LAST_X :	DWORD;
	END_VAR

	IF X > last_X THEN
		TU := TRUE;
		TD := FALSE;
		D := UDINT_TO_DWORD(DWORD_TO_UDINT(X) - DWORD_TO_UDINT(last_X));
		Q := TRUE;
	ELSIF X < last_X THEN
		TD := TRUE;
		TU := FALSE;
		D := UDINT_TO_DWORD(DWORD_TO_UDINT(last_X) - DWORD_TO_UDINT(X));
		Q := FALSE;
	ELSE
		TU := FALSE;
		TD := FALSE;
		D := DWORD#0;
	END_IF;
	last_X := X;
END_FUNCTION_BLOCK

FUNCTION_BLOCK _RMP_NEXT_Block
	VAR_INPUT
		E :	BOOL := TRUE;
		IN :	BYTE;
		TR :	TIME;
		TF :	TIME;
		TL :	TIME;
	END_VAR

	VAR_OUTPUT
		DIR :	BOOL;
		UP :	BOOL;
		DN :	BOOL;
	END_VAR

	VAR_IN_OUT
		OUT :	BYTE;
	END_VAR
	VAR
		rmx :	_RMP_B;
		dirx :	TREND_DW;
		t_lock :	TP;
		xen :	BOOL;
		xdir :	BOOL;
	END_VAR

	dirx(X := BYTE_TO_DWORD(in));

	t_lock(in := FALSE, pt := TL);

	IF dirx.TU AND (OUT < IN) THEN
		IF NOT xdir AND xen THEN t_lock(in := TRUE); END_IF;
		xen := TRUE;
		xdir := TRUE;
	ELSIF dirx.TD AND (OUT > IN) THEN
		IF xdir AND xen THEN t_lock(in := TRUE); END_IF;
		xen := TRUE;
		xdir := FALSE;
	ELSIF xen THEN
		IF (xdir AND (out >= in)) OR (NOT xdir AND (out <= in)) THEN
			xen := FALSE;
			IF tl > t#0s THEN t_lock(IN := TRUE); END_IF;
		END_IF;
	END_IF;

	IF NOT t_lock.Q AND xen THEN
		UP := XDIR;
		DIR := XDIR;
		DN := NOT XDIR;
	ELSE
		UP := FALSE;
		DN := FALSE;
	END_IF;

	rmx(rmp := OUT, E := E AND (UP OR DN) , dir := DIR, tr := SEL(dir, TF, TR));
	OUT := rmx.RMP;
END_FUNCTION_BLOCK

FUNCTION _BYTE_TO_INT:INT
	VAR_INPUT
		IN :	BYTE;
	END_VAR

	_BYTE_TO_INT := USINT_TO_INT(BYTE_TO_USINT(IN));
END_FUNCTION

FUNCTION_BLOCK ACTUATOR_3P_Block

	VAR_INPUT
		IN :	BYTE;
		TEST :	BOOL;
		ARE :	BOOL := TRUE;
		END_POS :	BOOL;
		T_RUN :	TIME := T#60s;
		T_EXT :	TIME := T#10s;
		T_CAL :	TIME := T#600s;
		T_DIAG :	TIME := T#10d;
		SWITCH_AVAIL :	BOOL;
	END_VAR

	VAR_OUTPUT
		OUT1 :	BOOL;
		OUT2 :	BOOL;
		POS :	BYTE;
		ERROR :	BOOL;
		STATUS :	BYTE;
	END_VAR

	VAR_IN_OUT
		ARX :	BOOL;
	END_VAR

	VAR
		tx :	TIME;
		_ramp :	_RMP_NEXT_Block;
		next_cal :	TIME;
		next_diag :	TIME;
		last :	TIME;
		start :	TIME;
		T_PLC_MS :	T_PLC_MS_Block;
	END_VAR

	T_PLC_MS();
	tx := UDINT_TO_TIME(T_PLC_MS.T_PLC_MS);

	IF TEST THEN
		status := BYTE#103;
		start := tx;
		ARX := TRUE;
	END_IF;

	CASE _BYTE_TO_INT(status) OF
		0:
			IF ARE AND NOT ARX THEN
				status := BYTE#103;
				start := tx;
				ARX := TRUE;
			END_IF;

		100:
			IF T_DIAG > T#0s AND tx > next_diag AND ARE AND NOT ARX THEN
					status := BYTE#103;
					start := tx;
					ARX := TRUE;

			ELSIF T_CAL > T#0s AND tx > next_cal AND ARE AND NOT ARX THEN
				IF pos > BYTE#127 THEN
					OUT1 := TRUE;
					OUT2 := FALSE;
					_ramp.IN := BYTE#255;
					ARX := TRUE;
				ELSE
					OUT1 := FALSE;
					OUT2 := TRUE;
					_ramp.IN := BYTE#0;
					ARX := TRUE;
				END_IF;
				status := BYTE#101;
				start := tx;
			ELSE
				IF NOT(OUT1 OR OUT2) THEN next_cal := next_cal + (tx-last); END_IF;
				_ramp.IN := IN;
			END_IF;

		101:
			IF tx - start < T_EXT THEN
				next_cal := tx + T_CAL;
			ELSIF SWITCH_AVAIL AND END_POS THEN
				STATUS := BYTE#100;
				ARX := FALSE;
			ELSIF tx - start > T_EXT + T_RUN THEN
				ERROR := SWITCH_AVAIL;
				ARX := FALSE;
			END_IF;

		103:
			IF tx - start < T_EXT THEN
				ERROR := FALSE;
				_ramp.TR := T_RUN;
				_ramp.TF := T_RUN;
				OUT1 := TRUE;
				OUT2 := FALSE;
				_ramp.IN := BYTE#255;
			ELSIF SWITCH_AVAIL AND END_POS THEN
				_ramp.TR := tx - start;
				STATUS := BYTE#104;
			ELSIF tx - start > T_EXT + T_RUN THEN
				ERROR := SWITCH_AVAIL;
				STATUS := BYTE#104;
				start := tx;
			END_IF;

		104:
			IF tx - start < T_ext THEN
				OUT1 := FALSE;
				OUT2 := TRUE;
				_ramp.IN := BYTE#0;
				next_diag := tx + T_DIAG;
			ELSIF SWITCH_AVAIL AND END_POS THEN
				_ramp.TR := tx - start;
				IF DINT_TO_TIME(ABS(TIME_TO_DINT(_ramp.TR) - TIME_TO_DINT(_ramp.TF)) * DINT#10) > T_RUN THEN error := TRUE; END_IF;
				STATUS := BYTE#100;
				ARX := FALSE;
				next_cal := tx + T_CAL;
			ELSIF tx - start > T_EXT + T_RUN THEN
				IF SWITCH_AVAIL THEN ERROR := TRUE; END_IF;
				STATUS := BYTE#100;
				ARX := FALSE;
				next_CAL := tx + T_CAL;
			END_IF;
	END_CASE;

	_ramp(OUT := POS);
	POS := _ramp.OUT;
	IF STATUS = BYTE#100 THEN
		OUT1 := _ramp.UP;
		OUT2 := _ramp.DN;
	END_IF;

	IF SWITCH_AVAIL AND END_POS THEN
		POS := SEL_BYTE(POS > BYTE#127, BYTE#0, BYTE#255);
		next_cal := tx + T_CAL;
	END_IF;

	last := tx;

END_FUNCTION_BLOCK

PROGRAM program0
	VAR
		IN :	BYTE;
		TEST :	BOOL;
		ARE :	BOOL := TRUE;
		END_POS :	BOOL;
		T_RUN :	TIME := T#60s;
		T_EXT :	TIME := T#10s;
		T_CAL :	TIME := T#600s;
		T_DIAG :	TIME := T#10d;
		SWITCH_AVAIL :	BOOL;
		OUT1 :	BOOL;
		OUT2 :	BOOL;
		POS :	BYTE;
		ERROR :	BOOL;
		STATUS :	BYTE;
		func_block : ACTUATOR_3P_Block;
	END_VAR
	func_block.IN := IN;
	func_block.TEST := TEST;
	func_block.ARE := ARE ;
	func_block.END_POS := END_POS;
	func_block.T_RUN := T_RUN;
	func_block.T_EXT := T_EXT;
	func_block.T_CAL := T_CAL ;
	func_block.T_DIAG := T_DIAG;
	func_block.SWITCH_AVAIL := SWITCH_AVAIL;
	func_block();
	OUT1  := func_block.OUT1;
	OUT2  := func_block.OUT2;
	POS  := func_block.POS;
	ERROR  := func_block.ERROR;
	STATUS  := func_block.STATUS;
END_PROGRAM

CONFIGURATION Config0
	VAR_GLOBAL
		PLC_TICKS_PER_SEC :	INT;
		PLC_SYS_TICK_CNT :	DINT;
	END_VAR
  	RESOURCE Res0 ON PLC
    	TASK task0(INTERVAL := T#20ms,PRIORITY := 0);
    	PROGRAM instance0 WITH task0 : program0;
  	END_RESOURCE
END_CONFIGURATION

(* ---- 724-BURNER.ST ---- *)
FUNCTION_BLOCK ONTIME_Block

	VAR_INPUT
		IN :	BOOL;
		RST :	BOOL;
	END_VAR

	VAR_IN_OUT
		SECONDS :	UDINT;
		CYCLES :	UDINT;
	END_VAR

	VAR
		tx :	UDINT;
		last :	UDINT;
		edge :	BOOL;
		init :	BOOL;
		ms :	UDINT;
		T_PLC_MS :	T_PLC_MS_Block;
	END_VAR

	T_PLC_MS();
	tx:= T_PLC_MS.T_PLC_MS;

	IF NOT init THEN
		init := TRUE;
		last := tx;
		ms := UDINT#0;
	END_IF;
	IF RST THEN
		SECONDS := UDINT#0;
		CYCLES := UDINT#0;
		last := tx;
		ms := UDINT#0;
	ELSIF IN THEN
		(* add the current milliseconds *)
		ms := (tx - last) + ms;
		IF ms >= UDINT#1000 THEN
			seconds := seconds + UDINT#1;
			ms := ms - UDINT#1000;
		END_IF;
		cycles := cycles + BOOL_TO_UDINT(NOT edge);
	END_IF;
	last := tx;
	edge := in;

END_FUNCTION_BLOCK

FUNCTION UDINT_TO_TIME2:TIME

	VAR_INPUT
		IN :	UDINT;
	END_VAR

	UDINT_TO_TIME2 := DINT_TO_TIME(UDINT_TO_DINT(IN));

END_FUNCTION

FUNCTION_BLOCK T_PLC_MS_block
	VAR_OUTPUT
		T_PLC_MS :	UDINT;
	END_VAR

	VAR_EXTERNAL
		PLC_TICKS_PER_SEC :	INT;
		PLC_SYS_TICK_CNT :	DINT;
	END_VAR

	VAR
		debug :	BOOL;(*Debug-Mode ON / OFF*)
		N :	INT;(*Debug-Faktor*)
		Offset :	UDINT;(*Debug-Offset*)
		temp :	DWORD := DWORD#1;(*Debug-Offset*)
		mode :	BOOL;(*modus*)
		faktor :	UDINT;(*Systemtakt-Faktor*)
		init :	BOOL;
		v_plc_ticks_per_sec :	UDINT;
		base :	UDINT := UDINT#1000;
	END_VAR

	IF init = FALSE THEN
		v_plc_ticks_per_sec := INT_TO_UDINT(PLC_TICKS_PER_SEC);
		IF v_plc_ticks_per_sec = UDINT#1024 THEN
			faktor := UDINT#1;
			mode := FALSE;
		ELSIF v_plc_ticks_per_sec > UDINT#0 THEN
			IF v_plc_ticks_per_sec <= base THEN
				faktor := base / v_plc_ticks_per_sec;
				mode := FALSE;
			ELSE
				faktor := v_plc_ticks_per_sec / base;
				mode := TRUE;
			END_IF;
		ELSE
			faktor := UDINT#1;
		END_IF;
		init := TRUE;
	END_IF;

	IF mode THEN
		T_PLC_MS := DINT_TO_UDINT(PLC_SYS_TICK_CNT) / faktor;
	ELSE
		T_PLC_MS := DINT_TO_UDINT(PLC_SYS_TICK_CNT) * faktor;
	END_IF;

	IF debug THEN
		T_PLC_MS := (DWORD_TO_UDINT(SHL(UDINT_TO_DWORD(T_PLC_MS),N) OR SHL(temp,N)) - UDINT#1) + Offset;
	END_IF;

END_FUNCTION_BLOCK

FUNCTION_BLOCK BURNER_Block

	VAR_INPUT
		IN :	BOOL;
		STAGE2 :	BOOL;
		OVER_TEMP :	BOOL;
		OIL_TEMP :	BOOL := TRUE;
		FLAME :	BOOL;
		RST :	BOOL;
		RST_TIMER :	BOOL;
		PRE_HEAT_TIME :	TIME := t#5s;
		PRE_VENT_TIME :	TIME := t#15s;
		PRE_IGNITE_TIME :	TIME := t#5s;
		POST_IGNITE_TIME :	TIME := t#25s;
		STAGE2_DELAY :	TIME := t#10s;
		SAFETY_TIME :	TIME := t#5s;
		LOCKOUT_TIME :	TIME := t#10s;
		MULTIPLE_IGNITION :	BOOL := TRUE;
		KW1 :	REAL;
		KW2 :	REAL;
	END_VAR

	VAR_OUTPUT
		MOTOR :	BOOL;
		COIL1 :	BOOL;
		COIL2 :	BOOL;
		PRE_HEAT :	BOOL;
		IGNITE :	BOOL;
		KWH :	REAL;
		STATUS :	BYTE;
		FAIL :	BOOL;
	END_VAR

	VAR_IN_OUT
		RUNTIME1 :	UDINT;
		RUNTIME2 :	UDINT;
		CYCLES :	UDINT;
	END_VAR

	VAR
		state :	INT;
		last :	TIME;
		tx :	TIME;
		last_change :	TIME;
		timer1 :	ONTIME_Block;
		timer2 :	ONTIME_Block;
		oil_temp_last :	BOOL;
		cycles2 :	UDINT;
		T_PLC_MS :	T_PLC_MS_Block;
	END_VAR

	T_PLC_MS();
	tx:= UDINT_TO_TIME(T_PLC_MS.T_PLC_MS);

	IF rst OR over_temp OR state = 0 THEN
		IF status > BYTE#0 AND tx - last_change >= lockout_time AND rst THEN
			status := BYTE#110;
			fail := FALSE;
			state := 1;
		ELSE
			motor := FALSE;
			coil1 := FALSE;
			coil2 := FALSE;
			ignite := FALSE;
			pre_heat := FALSE;
			IF over_temp THEN
				status := BYTE#9;
				fail := TRUE;
			END_IF;
			last_change := tx;
			last := tx;
			state := 1;
		END_IF;
	END_IF;

	IF rst_timer THEN
		runtime1 := UDINT#0;
		runtime2 := UDINT#0;
		cycles := UDINT#0;
		cycles2 := UDINT#0;
	END_IF;

	IF (status > BYTE#0 AND status < BYTE#100) OR rst THEN RETURN; END_IF;

	CASE state OF

	1:
		IF in AND flame THEN
			state := 7;
			pre_heat := FALSE;
			status := BYTE#2;
			last_change := tx;
		ELSIF in THEN
			pre_heat := TRUE;
			state := 2;
			last_change := tx;
		END_IF;

	2:
		IF (tx- last_change >= pre_heat_time AND oil_temp) OR (oil_temp AND NOT oil_temp_last) THEN
			motor := TRUE;
			state := 3;
			last_change := tx;
		ELSIF tx - last_change >= pre_heat_time AND NOT oil_temp THEN
			state := 7;
			pre_heat := FALSE;
			status := BYTE#1;
			last_change := tx;
		ELSIF flame THEN
			state := 7;
			pre_heat := FALSE;
			status := BYTE#2;
			last_change := tx;
		END_IF;

	3:
		IF tx - last_change >= pre_vent_time - pre_ignite_time THEN
			ignite := TRUE;
			state := 4;
			last_change := tx;
		ELSIF flame THEN
			state := 7;
			pre_heat := FALSE;
			motor := FALSE;
			status := BYTE#3;
			last_change := tx;
		END_IF;

	4:
		IF tx - last_change >= pre_ignite_time THEN
			coil1 := TRUE;
			state := 5;
			last_change := tx;
		END_IF;

	5:
		IF tx - last_change >= safety_time OR flame THEN
			IF NOT flame THEN
				state := 7;
				motor := FALSE;
				coil1 := FALSE;
				pre_heat := FALSE;
				ignite := FALSE;
				status := BYTE#4;
				last_change := tx;
			ELSE
				state := 6;
				last_change := tx;
			END_IF;
		END_IF;

	6:
		IF NOT flame AND NOT multiple_ignition THEN
			state := 7;
			motor := FALSE;
			coil1 := FALSE;
			coil2 := FALSE;
			pre_heat := FALSE;
			ignite := FALSE;
			status := BYTE#5;
			last_change := tx;
		ELSIF NOT flame AND multiple_ignition THEN
			ignite := TRUE;
			state := 5;
			coil2 := FALSE;
			last_change := tx;
		ELSE
			IF tx - last_change >= post_ignite_time THEN
				ignite := FALSE;
			END_IF;
			IF tx - last_change >= stage2_delay AND stage2 THEN
				coil2 := TRUE;
			ELSE
				coil2 := FALSE;
			END_IF;
		END_IF;
	END_CASE;

	IF NOT in THEN
		state := 1;
		motor := FALSE;
		coil1 := FALSE;
		coil2 := FALSE;
		ignite := FALSE;
		pre_heat := FALSE;
		last_change := tx;
	END_IF;

	timer1(in := flame AND in AND motor AND coil1 AND NOT coil2, SECONDS := runtime1, CYCLES := cycles);
	cycles := timer1.CYCLES;
	runtime1 := timer1.SECONDS;

	timer2(in := flame AND in AND motor AND coil1 AND coil2, SECONDS := runtime2, CYCLES := cycles2);
	cycles2 := timer2.CYCLES;
	runtime2 := timer2.SECONDS;

	KWH := UDINT_TO_REAL(runtime1) * KW1 / 3600.0 + UDINT_TO_REAL(runtime2) * KW2 / 3600.0;

	last := tx;

	IF status > BYTE#0 AND status < BYTE#100 THEN
		fail := TRUE;
	ELSE
		fail := FALSE;
		IF NOT in THEN
			status := BYTE#110;
		ELSIF flame AND in AND motor AND coil2 AND coil1 THEN
			status := BYTE#113;
		ELSIF flame AND in AND motor AND coil1 THEN
			status := BYTE#112;
		ELSE
			status := BYTE#111;
		END_IF;
	END_IF;

END_FUNCTION_BLOCK

PROGRAM program0
	VAR
		IN :	BOOL;
		STAGE2 :	BOOL;
		OVER_TEMP :	BOOL;
		OIL_TEMP :	BOOL := TRUE;
		FLAME :	BOOL;
		RST :	BOOL;
		RST_TIMER :	BOOL;
		PRE_HEAT_TIME :	TIME := t#5s;
		PRE_VENT_TIME :	TIME := t#15s;
		PRE_IGNITE_TIME :	TIME := t#5s;
		POST_IGNITE_TIME :	TIME := t#25s;
		STAGE2_DELAY :	TIME := t#10s;
		SAFETY_TIME :	TIME := t#5s;
		LOCKOUT_TIME :	TIME := t#10s;
		MULTIPLE_IGNITION :	BOOL := TRUE;
		KW1 :	REAL;
		KW2 :	REAL;
		RUNTIME1 :	UDINT;
		RUNTIME2 :	UDINT;
		CYCLES :	UDINT;
		MOTOR :	BOOL;
		COIL1 :	BOOL;
		COIL2 :	BOOL;
		PRE_HEAT :	BOOL;
		IGNITE :	BOOL;
		KWH :	REAL;
		STATUS :	BYTE;
		FAIL :	BOOL;

		func_block : BURNER_Block;
	END_VAR
	func_block.IN := IN;
	func_block.STAGE2 := STAGE2;
	func_block.OVER_TEMP := OVER_TEMP ;
	func_block.OIL_TEMP    := OIL_TEMP    ;
	func_block.FLAME := FLAME;
	func_block.RST := RST;
	func_block.RST_TIMER := RST_TIMER ;
	func_block.PRE_HEAT_TIME := PRE_HEAT_TIME ;
	func_block.PRE_VENT_TIME    := PRE_VENT_TIME    ;
	func_block.PRE_IGNITE_TIME := PRE_IGNITE_TIME;
	func_block.POST_IGNITE_TIME := POST_IGNITE_TIME;
	func_block.STAGE2_DELAY := STAGE2_DELAY ;
	func_block.SAFETY_TIME := SAFETY_TIME ;
	func_block.LOCKOUT_TIME    := LOCKOUT_TIME    ;
	func_block.MULTIPLE_IGNITION := MULTIPLE_IGNITION;
	func_block.KW1 := KW1;
	func_block.KW2 := KW2;
	func_block.RUNTIME1 := RUNTIME1;
	func_block.RUNTIME2 := RUNTIME2;
	func_block.CYCLES := CYCLES;

	func_block();
	MOTOR  := func_block.MOTOR;
	COIL1  := func_block.COIL1;
	COIL2  := func_block.COIL2;
	PRE_HEAT  := func_block.PRE_HEAT;
	IGNITE  := func_block.IGNITE;
	KWH  := func_block.KWH;
	STATUS  := func_block.STATUS;
	FAIL  := func_block.FAIL;
	RUNTIME1  := func_block.RUNTIME1;
	RUNTIME2  := func_block.RUNTIME2;
	CYCLES  := func_block.CYCLES;
END_PROGRAM

CONFIGURATION Config0
	VAR_GLOBAL
		PLC_TICKS_PER_SEC :	INT;
		PLC_SYS_TICK_CNT :	DINT;
	END_VAR
  	RESOURCE Res0 ON PLC
    	TASK task0(INTERVAL := T#20ms,PRIORITY := 0);
    	PROGRAM instance0 WITH task0 : program0;
  	END_RESOURCE
END_CONFIGURATION

(* ---- 725-IP_CONTROL.ST ---- *)
FUNCTION_BLOCK IP_CONTROL_Block

  VAR
    T_PLC_MS :	T_PLC_MS;
    IP4_TO_STRING :	IP4_TO_STRING;
    FB_IP_CONNECT :	IP_CONNECT;
    FB_IP_URCV :	IP_URCV;
    FB_IP_USEND :	IP_USEND;
  END_VAR

  VAR_INPUT
    IP :	DWORD;
    PORT :	WORD;
    TIME_OUT :	TIME;
  END_VAR

  VAR_IN_OUT
    IP_C :	oscat_IP_C;
    S_BUF :	oscat_NETWORK_BUFFER;
    R_BUF :	oscat_NETWORK_BUFFER;
  END_VAR

  VAR
    C_TIME :	UDINT;
    S_TIME :	UDINT;
    R_TIME :	UDINT;
    C_ENABLE :	BOOL;
    C_IP :	DWORD;
    C_PORT :	WORD;
    C_MODE :	BYTE;
    C_ERROR :	BOOL;
    C_STATUS :	INT;
    C_ID :	INT;
    C_RECONNECT :	BOOL;
    C_RECONNECT_COUNT :	INT;
    S_BUF_I :	oscat_NETWORK_BUFFER_SHORT;
    S_TOTAL :	INT;
    S_CUR_POS :	INT;
    S_CUR_SIZE :	INT;
    S_MAX_SIZE :	INT := 1408;
    S_START :	BOOL;
    S_REQ :	BOOL;
    S_DONE :	BOOL;
    S_ERROR :	BOOL;
    S_STATUS :	INT;
    R_NDR :	BOOL;
    R_ERROR :	BOOL;
    R_STATUS :	INT;
    R_BUF_I :	oscat_NETWORK_BUFFER_SHORT;
    R_COUNT :	INT;
    R_OFFSET :	INT;
    R_E_MAX_SIZE :	INT := 4096;
    NEW_CONNECTION :	BOOL;
    C_ENABLE_OLD :	BOOL;
    C_READY :	BOOL;
    C_READY_OLD :	BOOL;
    DELAY_STOP :	UDINT;
    DELAY :	UDINT;
    DELAY_VALUE :	UDINT;
    C :	INT;
    C2 :	INT;
    C3 :	INT;
    CS :	STRING;
    TX :	UDINT;
    ERROR_TIME :	UDINT;
    S_ACTIVE :	BOOL;
    ERROR_CON :	BYTE;
    ERROR_SND :	BYTE;
    ERROR_RCV :	BYTE;
  END_VAR

  T_PLC_MS();
  TX := T_PLC_MS.T_PLC_MS;

  IF (TX - DELAY < DELAY_VALUE) THEN
    IF IP_C.C_STATE <> BYTE#1 AND IP_C.C_STATE <> BYTE#254 THEN
    RETURN;
    END_IF;
  END_IF;
  DELAY := TX;

  IF C_ENABLE AND DELAY_VALUE > UDINT#00 THEN
    IF (TX - DELAY_STOP > UDINT#1000) THEN
      DELAY_VALUE := UDINT#00;
    END_IF;
  ELSE
    DELAY_STOP := TX;
  END_IF;

  IF IP_C.C_PORT = WORD#00 THEN
    IP_C.C_PORT := PORT;
  END_IF;
  IF IP_C.C_IP=DWORD#00 AND IP_C.C_MODE<BYTE#4 THEN
    IP_C.C_IP := IP;
  END_IF;

  NEW_CONNECTION := C_IP <> IP_C.C_IP OR C_MODE <> IP_C.C_MODE OR C_PORT <> IP_C.C_PORT;

  IF IP_C.C_ENABLE AND NOT C_READY AND NEW_CONNECTION THEN

    C_IP   := IP_C.C_IP;
    C_MODE := IP_C.C_MODE;
    C_PORT := IP_C.C_PORT;

    CS := SEL_STRING((C_MODE AND BYTE#1) = BYTE#1,'','/UDP');
    CS := CONCAT(CS,SEL_STRING(C_MODE<BYTE#2,' /PASSIVE',' /ACTIVE'));
    CS := CONCAT(CS,' /PORT=');
    CS := CONCAT(CS,WORD_TO_STRING(C_PORT,'%u'));

    IF C_MODE<BYTE#4 THEN
      IP4_TO_STRING(IP4:=C_IP);
      CS := CONCAT(CS,' /IP=');
      CS := CONCAT(CS,IP4_TO_STRING.IP4_TO_STRING);
    END_IF;

    ERROR_TIME := MAX(UDINT#200,TIME_TO_UDINT2(TIME_OUT));
    IP_C.TIME_RESET := TRUE;
  END_IF;

  C_ENABLE := IP_C.C_ENABLE AND NOT C_RECONNECT AND NOT NEW_CONNECTION AND IP_C.ERROR = DWORD#0;

  FB_IP_CONNECT.EN_C    := C_ENABLE;
  FB_IP_CONNECT.PARTNER := CS;
  FB_IP_CONNECT();
  C_READY  := FB_IP_CONNECT.VALID;
  C_ERROR  := FB_IP_CONNECT.ERROR;
  C_STATUS := FB_IP_CONNECT.STATUS;
  C_ID     := FB_IP_CONNECT.ID;

  IF C_ENABLE THEN
    IF NOT C_ENABLE_OLD THEN
      DELAY_VALUE := UDINT#50;
    END_IF;
  ELSE
    IF C_ENABLE_OLD THEN
      C_RECONNECT := FALSE;
      DELAY_VALUE := UDINT#50;
    END_IF;
  END_IF;

  C_ENABLE_OLD := C_ENABLE;

  IF C_READY THEN
    IF NOT C_READY_OLD THEN
      IP_C.C_STATE := BYTE#254;
      DELAY_VALUE := UDINT#50;
      IP_C.TIME_RESET := TRUE;

    ELSE
      IP_C.C_STATE := BYTE#255;
    END_IF;
  ELSE
    IF C_READY_OLD THEN
      IP_C.C_STATE := BYTE#1;
    IP_C.MAILBOX[1] := BYTE#0;
    IP_C.MAILBOX[2] := BYTE#0;
    IP_C.MAILBOX[3] := BYTE#0;
      DELAY_VALUE := UDINT#50;

      IF NOT NEW_CONNECTION THEN
        S_ACTIVE := FALSE;
        S_REQ := FALSE;
        S_BUF.SIZE := UINT#0;
      END_IF;
    ELSE
      IP_C.C_STATE := BYTE#000;
    END_IF;
  END_IF;

  C_READY_OLD := C_READY;

  C := 1;
  IF S_BUF.SIZE > UINT#0 THEN
    IF C_READY AND C_ENABLE THEN
      IF S_ACTIVE = FALSE AND IP_C.MAILBOX[2] = BYTE#0 THEN
        S_TOTAL := LIMIT_INT(0,UINT_TO_INT(S_BUF.SIZE),R_E_MAX_SIZE);
        S_CUR_POS  := 0;
        S_CUR_SIZE := 0;
        S_START := TRUE;
        S_ACTIVE := TRUE;
      END_IF;

      IF S_DONE OR S_START THEN

        S_START := FALSE;
        S_CUR_POS := S_CUR_POS + S_CUR_SIZE;
        IF S_TOTAL > S_CUR_POS THEN
          S_CUR_SIZE := S_TOTAL - S_CUR_POS;
          S_CUR_SIZE:=LIMIT_INT(0,S_CUR_SIZE,S_MAX_SIZE);

          C2 := S_CUR_POS;
      C3 := S_CUR_SIZE - 1;
      FOR C := 0 TO C3 DO
            S_BUF_I.BUFFER[C] := S_BUF.BUFFER[C2];
        C2 := C2 + 1;
          END_FOR;
          S_BUF_I.SIZE := INT_TO_UINT(S_CUR_SIZE);
        S_TIME := tx;
          R_TIME := tx;
          S_REQ := TRUE;
          C := 0;
        ELSE
          S_REQ := FALSE;
          S_BUF.SIZE := UINT#0;
          S_ACTIVE := FALSE;
        END_IF;
      END_IF;
    END_IF;
  END_IF;

  FOR C2 := C TO 1 DO
    FB_IP_USEND.REQ    := S_REQ AND C2=1;
    FB_IP_USEND.ID     := C_ID;
    FB_IP_USEND.R_ID   := '';
    FB_IP_USEND.SD_1   := S_BUF_I;
    FB_IP_USEND();
    S_DONE   := FB_IP_USEND.DONE;
    S_ERROR  := FB_IP_USEND.ERROR;
    S_STATUS := FB_IP_USEND.STATUS;
    S_BUF_I  := FB_IP_USEND.SD_1;
  END_FOR;

  FB_IP_URCV.EN_R := C_READY AND NOT S_ACTIVE AND IP_C.MAILBOX[3] = BYTE#0;
  FB_IP_URCV.ID   := C_ID;
  FB_IP_URCV.R_ID := '';
  FB_IP_URCV.RD_1 := R_BUF_I;
  FB_IP_URCV();
  R_NDR    := FB_IP_URCV.NDR;
  R_ERROR  := FB_IP_URCV.ERROR;
  R_STATUS := FB_IP_URCV.STATUS;
  R_BUF_I  := FB_IP_URCV.RD_1;

  IF R_NDR THEN
    IF R_BUF.SIZE >= INT_TO_UINT(R_E_MAX_SIZE) THEN
      R_BUF.SIZE := UINT#0;
      r_status := 254;
    END_IF;

    R_TIME := tx;
    R_COUNT := UINT_TO_INT(R_BUF_I.SIZE);
    R_OFFSET := UINT_TO_INT(R_BUF.SIZE);

    IF (C_MODE AND BYTE#2#0000_0001) = BYTE#1 THEN
      r_offset := 0;
    ELSE
      R_OFFSET := UINT_TO_INT(R_BUF.SIZE);
    END_IF;

    IF R_OFFSET + R_COUNT > R_E_MAX_SIZE THEN
      R_COUNT := R_E_MAX_SIZE - R_OFFSET;
    END_IF;

    C2 := R_OFFSET;
    C3 := R_COUNT - 1;
    FOR C := 0 TO C3 DO
      R_BUF.BUFFER[C2] := R_BUF_I.BUFFER[C];
      C2 := C2 + 1;
    END_FOR;

    R_BUF.SIZE := INT_TO_UINT(R_OFFSET + R_COUNT);
    IP_C.MAILBOX[1] := USINT_TO_BYTE(BYTE_TO_USINT(IP_C.MAILBOX[1]) + USINT#1);
    IF IP_C.MAILBOX[1] = BYTE#0 THEN IP_C.MAILBOX[1] := BYTE#1; END_IF;

  END_IF;

  IF IP_C.TIME_RESET THEN
    IP_C.TIME_RESET := FALSE;
    C_RECONNECT_COUNT := 0;
    C_TIME := tx;
    S_TIME := tx;
    R_TIME := tx;

    ERROR_CON := BYTE#0;
    ERROR_SND := BYTE#0;
    ERROR_RCV := BYTE#0;
  END_IF;

  IF IP_C.R_OBSERVE = FALSE OR s_active THEN
      R_TIME := tx;
  END_IF;

  C_RECONNECT := FALSE;

  IF ERROR_CON = BYTE#0 THEN
    IF C_ERROR THEN
    IF C_STATUS = 16#31 THEN
      ERROR_CON := BYTE#253;
    ELSE
      ERROR_CON := INT_TO_BYTE(C_STATUS);
    END_IF;
    ELSIF TX - C_TIME > ERROR_TIME AND C_ENABLE AND NOT C_READY AND C_MODE < BYTE#2 THEN
      IF C_RECONNECT_COUNT >= 3 THEN
        ERROR_CON := BYTE#255;
      ELSE
        C_TIME := TX;
        C_RECONNECT_COUNT := C_RECONNECT_COUNT + 1;
        C_RECONNECT := TRUE;

      END_IF;
    END_IF;
  END_IF;

  IF ERROR_SND = BYTE#0 THEN
    IF S_ERROR AND S_STATUS <> 16#65 THEN
      ERROR_SND := INT_TO_BYTE(S_STATUS);
    ELSIF TX - S_TIME > ERROR_TIME AND S_ACTIVE THEN
      ERROR_SND := BYTE#255;
    END_IF;
  END_IF;

  IF ERROR_RCV = BYTE#0 THEN
    IF R_ERROR AND (R_STATUS <> 16#33) AND (R_STATUS <> 16#31) AND (R_STATUS <> 16#65) THEN
      ERROR_RCV := INT_TO_BYTE(R_STATUS);
    ELSIF TX - R_TIME > ERROR_TIME AND C_READY AND IP_C.R_OBSERVE THEN
      ERROR_RCV := BYTE#255;
    END_IF;
  END_IF;

  IP_C.ERROR := DWORD_OF_BYTE(ERROR_CON,ERROR_SND,ERROR_RCV,BYTE#0);

END_FUNCTION_BLOCK

PROGRAM program0
	VAR
		IP :	DWORD;
    PORT :	WORD;
    TIME_OUT :	TIME;
    IP_C :	oscat_IP_C;
    S_BUF :	oscat_NETWORK_BUFFER;
    R_BUF :	oscat_NETWORK_BUFFER;

		func_block : IP_CONTROL_Block;
	END_VAR
	func_block.IP := IP;
	func_block.PORT := PORT;
	func_block.TIME_OUT := TIME_OUT;
	func_block.IP_C := IP_C;
	func_block.S_BUF := S_BUF;
	func_block.R_BUF := R_BUF;

	func_block();
  IP_C  := func_block.IP_C;
	S_BUF  := func_block.S_BUF;
	R_BUF  := func_block.R_BUF;

END_PROGRAM

CONFIGURATION Config0
	RESOURCE Res0 ON PLC
		TASK task0(INTERVAL := T#20ms,PRIORITY := 0);
		PROGRAM instance0 WITH task0 : program0;
	END_RESOURCE
END_CONFIGURATION

(* ---- 726-SNTP_SERVER.ST ---- *)
TYPE
  oscat_IP_FIFO128_DATA  : ARRAY [1..128] OF BYTE;
  oscat_Mailbox  : ARRAY [1..16] OF BYTE;

  oscat_IP_FIFO_DATA :
  STRUCT
    X       : oscat_IP_FIFO128_DATA; (* IP_ID FIFO Speicher          *)
    Y       : oscat_IP_FIFO128_DATA; (* IP_ID Z�hler                 *)
    ID      : BYTE;                  (* h�chste vergabene id         *)
    MAX_ID  : BYTE;                  (* maximal Anmeldungen pro ID   *)
      INIT    : BOOL;                  (* Initialisierung durchgef�hrt *)
    EMPTY   : BOOL;                  (* FIFO leer                    *)
    FULL    : BOOL;                  (* FIFO voll                    *)
    TOP     : INT;                   (* maximale anzahl in FIFO      *)
    NW      : INT;                   (* Schreibzeiger                *)
    NR      : INT;                   (* Lesezeiger                   *)
  END_STRUCT;

  oscat_IP_C:
  STRUCT
    C_MODE:			BYTE;          		(*W Mode: TCP/UCP AKTIV/PASSIV                               *)
    C_PORT:         WORD;          		(*W Portnummer                                               *)
    C_IP:           DWORD;         		(*W IP-Adresse gepackt wwxxyyzz = www.xxx.yyy.zzz            *)
    C_STATE:        BYTE;          		(*R Verbindungsstatus ON/OFF + Flanke ON/OFF                 *)
    C_ENABLE:       BOOL;          		(*W Freigabe f�r Connect                                     *)
    R_OBSERVE:      BOOL;          		(*W Empfang ueberwachen                                      *)
    TIME_RESET:     BOOL;          		(*W Alle Timer ruecksetzen                                   *)
    ERROR:          DWORD;         		(*R vvwwxxyy (vv = CON_ERROR, ww = SEN_ERROR, xx = REC_ERROR *)
    FIFO:           oscat_IP_FIFO_DATA; (*I IP FIFO Struktur                                         *)
    MAILBOX:		oscat_Mailbox;		(*I Mailbox: Datenbereich f�r Bausteindatenaustausch         *)
  END_STRUCT;
END_TYPE

TYPE

  oscat_NW_BUF_LONG  : ARRAY [0..4095] OF BYTE;

  oscat_NETWORK_BUFFER :
  STRUCT
    SIZE   : UINT;
    BUFFER : oscat_NW_BUF_LONG;
  END_STRUCT;

END_TYPE

FUNCTION _BYTE_TO_INT:INT
	VAR_INPUT
		IN :	BYTE;
	END_VAR

	_BYTE_TO_INT := USINT_TO_INT(BYTE_TO_USINT(IN));
END_FUNCTION

FUNCTION_BLOCK IP_FIFO_Block

  VAR_IN_OUT
    FIFO :	oscat_IP_FIFO_DATA;
    ID :	BYTE;
    STATE :	BYTE;
  END_VAR

  VAR
    tmp :	INT;
  END_VAR

  IF NOT FIFO.INIT THEN
    FIFO.INIT		:= TRUE;
    FIFO.NW		:= 1;
    FIFO.NR		:= 1;
    FIFO.EMPTY	:= TRUE;
    FIFO.FULL		:= FALSE;
    FIFO.TOP		:= 128;
    FIFO.MAX_ID	:= BYTE#1;
  END_IF;

  IF ID = BYTE#00 THEN
    IF FIFO.ID < INT_TO_BYTE(FIFO.TOP) THEN
      ID := USINT_TO_BYTE(BYTE_TO_USINT(FIFO.ID) + USINT#1);
      FIFO.ID := ID ;

    ELSIF STATE < BYTE#200 THEN
      STATE := BYTE#255;
    RETURN;
    END_IF;
  END_IF;

  IF STATE = BYTE#1 AND NOT FIFO.FULL THEN
    tmp := _BYTE_TO_INT(ID);
    IF FIFO.Y[tmp] < FIFO.MAX_ID THEN
      FIFO.Y[tmp] := USINT_TO_BYTE(BYTE_TO_USINT(FIFO.Y[tmp]) + USINT#1);
      tmp := FIFO.NW;
      FIFO.X[tmp] := ID;
      IF FIFO.NW = FIFO.TOP THEN FIFO.NW := 1; ELSE FIFO.NW := FIFO.NW + 1; END_IF;
      FIFO.FULL := FIFO.NW = FIFO.NR;
    FIFO.EMPTY := FALSE;
      STATE := BYTE#2;
    END_IF;
  END_IF;

  IF STATE = BYTE#2 AND NOT FIFO.EMPTY THEN
    tmp := FIFO.NR;
    IF ID = FIFO.X[tmp] THEN
      STATE := BYTE#3;
    END_IF;
  END_IF;

  IF STATE = BYTE#4 AND NOT FIFO.EMPTY THEN

    tmp := FIFO.NR;
    IF ID = FIFO.X[tmp] THEN
      tmp := _BYTE_TO_INT(ID);
      FIFO.Y[tmp] := USINT_TO_BYTE(BYTE_TO_USINT(FIFO.Y[tmp]) - USINT#1);

      IF FIFO.NR = FIFO.TOP THEN FIFO.NR := 1; ELSE FIFO.NR := FIFO.NR + 1; END_IF;
      FIFO.EMPTY := FIFO.NR = FIFO.NW;
    FIFO.FULL := FALSE;
    END_IF;
    STATE := BYTE#5;
  END_IF;

END_FUNCTION_BLOCK

FUNCTION_BLOCK T_PLC_MS_block

	VAR_OUTPUT
		T_PLC_MS :	UDINT;
	END_VAR

	VAR_EXTERNAL
		PLC_TICKS_PER_SEC :	INT;
		PLC_SYS_TICK_CNT :	DINT;
	END_VAR

	VAR
		debug :	BOOL;(*Debug-Mode ON / OFF*)
		N :	INT;(*Debug-Faktor*)
		Offset :	UDINT;(*Debug-Offset*)
		temp :	DWORD := DWORD#1;(*Debug-Offset*)
		mode :	BOOL;(*modus*)
		faktor :	UDINT;(*Systemtakt-Faktor*)
		init :	BOOL;
		v_plc_ticks_per_sec :	UDINT;
		base :	UDINT := UDINT#1000;
	END_VAR

	IF init = FALSE THEN
		v_plc_ticks_per_sec := INT_TO_UDINT(PLC_TICKS_PER_SEC);
		IF v_plc_ticks_per_sec = UDINT#1024 THEN
			faktor := UDINT#1;
			mode := FALSE;
		ELSIF v_plc_ticks_per_sec > UDINT#0 THEN
			IF v_plc_ticks_per_sec <= base THEN
				faktor := base / v_plc_ticks_per_sec;
				mode := FALSE;
			ELSE
				faktor := v_plc_ticks_per_sec / base;
				mode := TRUE;
			END_IF;
		ELSE
			faktor := UDINT#1;
		END_IF;
		init := TRUE;
	END_IF;

	IF mode THEN
		T_PLC_MS := DINT_TO_UDINT(PLC_SYS_TICK_CNT) / faktor;
	ELSE
		T_PLC_MS := DINT_TO_UDINT(PLC_SYS_TICK_CNT) * faktor;
	END_IF;

	IF debug THEN
		T_PLC_MS := (DWORD_TO_UDINT(SHL(UDINT_TO_DWORD(T_PLC_MS),N) OR SHL(temp,N)) - UDINT#1) + Offset;
	END_IF;

END_FUNCTION_BLOCK

FUNCTION_BLOCK SNTP_SERVER_Block

  VAR_IN_OUT
    IP_C :	oscat_IP_C;
    S_BUF :	oscat_NETWORK_BUFFER;
    R_BUF :	oscat_NETWORK_BUFFER;
  END_VAR

  VAR_INPUT
    ENABLE :	BOOL;
    STRATUM :	BYTE := BYTE#1;
    UDT :	UDINT;
    XMS :	INT;
  END_VAR

  VAR
    IP_STATE :	BYTE;
    IP_ID :	BYTE;
    IP_FIFO :	IP_FIFO_Block;
    i2 :	INT;
    i :	INT;
    TIMESTAMP_INT :	DWORD;
    TIMESTAMP_SEK :	DWORD;
    TS_B :	BYTE;
    state :	INT;
    T_PLC_MS :	T_PLC_MS_Block;
    tx :	UDINT;
    t :	TON;
  END_VAR

  T_PLC_MS();
  tx := T_PLC_MS.T_PLC_MS;

  CASE state OF

  00:
    IF ENABLE THEN
      state := 10;
      IP_STATE := BYTE#1;
    END_IF;

  10:
    IF IP_STATE = BYTE#3 THEN

      IP_C.C_PORT     := WORD#123;
      IP_C.C_IP       := DWORD#00;
      IP_C.C_MODE     := BYTE#5;
      IP_C.C_ENABLE   := TRUE;
      IP_C.TIME_RESET := TRUE;
      IP_C.R_OBSERVE  := FALSE;
      S_BUF.SIZE      := UINT#0;
      R_BUF.SIZE      := UINT#0;

      state := 20;
    END_IF;

  20:
    IF R_BUF.SIZE > UINT#0 THEN
      state := 20;
      FOR i := 0 TO 47 DO
        IF INT_TO_UINT(i) > R_BUF.SIZE - UINT#1 THEN
          R_BUF.BUFFER[i] := BYTE#00;
      END_IF;
        S_BUF.BUFFER[i] := BYTE#00;
      END_FOR;

    R_BUF.SIZE := UINT#0;

      S_BUF.BUFFER[0] := BYTE#2#11100;
      S_BUF.BUFFER[1] := STRATUM;
      S_BUF.BUFFER[2] := BYTE#10;
      S_BUF.BUFFER[3] := BYTE#16#FB;

      TIMESTAMP_INT := UDINT_TO_DWORD(UDT + UDINT#2208988800);

    TIMESTAMP_SEK := DINT_TO_DWORD(DWORD_TO_DINT(SHL(INT_TO_DWORD(XMS),16))/DINT#1000);

      TS_B := TIMESTAMP_INT.B3;
      S_BUF.BUFFER[16] := TS_B;
      S_BUF.BUFFER[32] := TS_B;
      S_BUF.BUFFER[40] := TS_B;

      TS_B := TIMESTAMP_INT.B2;
      S_BUF.BUFFER[17] := TS_B;
      S_BUF.BUFFER[33] := TS_B;
      S_BUF.BUFFER[41] := TS_B;

      TS_B := TIMESTAMP_INT.B1;
      S_BUF.BUFFER[18] := TS_B;
      S_BUF.BUFFER[34] := TS_B;
      S_BUF.BUFFER[42] := TS_B;

      TS_B := TIMESTAMP_INT.B0;
      S_BUF.BUFFER[19] := TS_B;
      S_BUF.BUFFER[35] := TS_B;
      S_BUF.BUFFER[43] := TS_B;

      TS_B := TIMESTAMP_SEK.B1;
      S_BUF.BUFFER[20] := TS_B;
      S_BUF.BUFFER[36] := TS_B;
      S_BUF.BUFFER[44] := TS_B;

      TS_B := TIMESTAMP_SEK.B0;
      S_BUF.BUFFER[21] := TS_B;
      S_BUF.BUFFER[37] := TS_B;
      S_BUF.BUFFER[45] := TS_B;

      i2 := 40;
      FOR i := 24 TO 31 DO
        S_BUF.BUFFER[i] := R_BUF.BUFFER[i2];
        i2 := i2 +1;
      END_FOR;

      S_BUF.SIZE := UINT#48;

    ELSIF NOT ENABLE AND S_BUF.SIZE = UINT#0 THEN
      IP_STATE := BYTE#4;
      state := 0;
    END_IF;

  END_CASE;

  t(IN:= IP_C.ERROR > DWORD#0, PT:=T#5s);
  IF t.Q THEN
    IP_C.TIME_RESET := TRUE;
  END_IF;

  IP_FIFO(FIFO:=IP_C.FIFO,STATE:=IP_STATE,ID:=IP_ID);
  IP_C.FIFO:=IP_FIFO.FIFO;
  IP_STATE := IP_FIFO.STATE;
  IP_ID:=IP_FIFO.ID;

END_FUNCTION_BLOCK

PROGRAM program0
	VAR
		IP_C :	oscat_IP_C;
    S_BUF :	oscat_NETWORK_BUFFER;
    R_BUF :	oscat_NETWORK_BUFFER;
    ENABLE :	BOOL;
    STRATUM :	BYTE := BYTE#1;
    UDT :	UDINT;
    XMS :	INT;

		func_block : SNTP_SERVER_Block;
	END_VAR
	func_block.IP_C := IP_C;
	func_block.S_BUF := S_BUF;
	func_block.R_BUF := R_BUF;
  func_block.ENABLE := ENABLE;
	func_block.STRATUM := STRATUM;
	func_block.UDT := UDT;
  func_block.XMS := XMS;

	func_block();
  IP_C  := func_block.IP_C;
  S_BUF  := func_block.S_BUF;
  R_BUF  := func_block.R_BUF;
END_PROGRAM

CONFIGURATION Config0

	VAR_GLOBAL
		PLC_TICKS_PER_SEC :	INT;
		PLC_SYS_TICK_CNT :	DINT;
	END_VAR

  	RESOURCE Res0 ON PLC
    	TASK task0(INTERVAL := T#20ms,PRIORITY := 0);
    	PROGRAM instance0 WITH task0 : program0;
  	END_RESOURCE

END_CONFIGURATION
